(* IEC 61131-3 sources: TetherPLC/tests/compat (part 3) *)

(* ---- tc2_ncfifoaxes_case.st ---- *)
PROGRAM Tc2NciFifoCase
VAR
    mask   AT %QD0 : DINT;
    st     : INT;
    prevSt : INT;
    cur    : INT;
    pulse  : BOOL;
    ax     : FB_MotionAxis;
    axM    : UDINT;
    axS    : UDINT;
    pwrM   : MC_Power;
    pwrS   : MC_Power;
    integ1 : FiFoGroupIntegrate;
    integ2 : FiFoGroupIntegrate;
    dim    : FiFoGetDimension;
    wr     : FiFoWrite;
    owr    : FiFoOverwrite;
    ovr    : FiFoSetChannelOverride;
    start  : FiFoStart;
    dis    : FiFoGroupDisintegrate;
    mon    : FB_Fifo;
    dim2   : FiFoGetDimension;
    rpM    : MC_ReadActualPosition;
    rpS    : MC_ReadActualPosition;
    data   : ARRAY[0..255] OF LREAL;
    k      : UDINT;
    enSig  : BOOL;
    finishedSeen : BOOL;
    seqOk  : BOOL;
    seqOk2 : BOOL;
    posOk1 : BOOL;
    posOk2 : BOOL;
    startEx : BOOL;
END_VAR

// Stage machine: one stage per scan via the cur snapshot.
cur := st;
IF cur <> prevSt THEN pulse := TRUE; ELSE pulse := FALSE; END_IF;
prevSt := cur;

// Channel monitor: status+poll every scan. In-process backends
// consume one queued row per poll; the IO backend consumes rows on
// the mc.time drive clock (poll is a no-op there).
mon.OP := 6;
mon.CHAN := 0;
mon();

enSig := (st >= 1) AND (st <= 40);
// FiFoStart is invoked every scan so its Execute edge tracking stays
// live across the two run stages.
startEx := pulse AND ((cur = 6) OR (cur = 10));
start(bExecute := startEx, iChannelId := 0, tTimeout := T#1S);
pwrM(Enable := enSig, Enable_Positive := TRUE, Enable_Negative := TRUE,
    Axis := axM);
pwrS(Enable := enSig, Enable_Positive := TRUE, Enable_Negative := TRUE,
    Axis := axS);
rpM(Enable := TRUE, Axis := axM);
rpS(Enable := TRUE, Axis := axS);

IF cur = 0 THEN
    ax.UNITS_PER_REV := 1000;
    ax.MAX_VEL := 2000;
    ax.MAX_ACCEL := 8000;
    ax.MAX_DECEL := 8000;
    ax.POS_MIN := -200000;
    ax.POS_MAX := 200000;
    ax.HOME_OFFSET := 0;
    ax.FOLLOW_WINDOW := 3;
    ax.FLAGS := 1;
    ax.OP := 1; ax();
    IF ax.AXIS <> 0 THEN axM := ax.AXIS; END_IF;
    ax.OP := 1; ax();
    IF ax.AXIS <> 0 THEN axS := ax.AXIS; END_IF;
    IF axM <> 0 AND axS <> 0 THEN
        mask := mask + 1;                       // bit0: two axes
        st := 1;
    END_IF;
ELSIF cur = 1 THEN
    IF pwrM.Status AND pwrS.Status THEN
        mask := mask + 2;                       // bit1: powered
        st := 2;
    END_IF;
ELSIF cur = 2 THEN
    integ1(bExecute := pulse, iChannelId := 0, iAxisId := axM,
           iGroupPosition := 1, tTimeout := T#1S);
    integ2(bExecute := pulse, iChannelId := 0, iAxisId := axS,
           iGroupPosition := 2, tTimeout := T#1S);
    IF pulse AND NOT integ1.bError AND NOT integ2.bError THEN
        mask := mask + 4;                       // bit2: integrated
        st := 3;
    END_IF;
ELSIF cur = 3 THEN
    dim(bExecute := pulse, iChannelId := 0, tTimeout := T#1S);
    IF dim.bError = FALSE THEN
        IF dim.iAxes = 2 AND dim.iMaxRows >= 100 THEN
            mask := mask + 8;                   // bit3: dimension
            st := 4;
        END_IF;
    END_IF;
ELSIF cur = 4 THEN
    // two rows x two axes: [100,200] then [300,400]
    data[0] := 100.0; data[1] := 200.0;
    data[8] := 300.0; data[9] := 400.0;
    wr(bExecute := pulse, iChannelId := 0,
       AdrDataArray := data, iRowsToWrite := 2, tTimeout := T#1S);
    IF pulse AND NOT wr.bError THEN
        mask := mask + 16;                      // bit4: write
        st := 5;
    END_IF;
ELSIF cur = 5 THEN
    ovr(bExecute := pulse, iChannelId := 0, iOverride := 150,
        tTimeout := T#1S);
    IF pulse AND NOT ovr.bError THEN
        mask := mask + 32;                      // bit5: override
        st := 6;
    END_IF;
ELSIF cur = 6 THEN
    IF pulse AND NOT start.bError THEN
        mask := mask + 64;                      // bit6: start
        st := 7;
    END_IF;
ELSIF cur = 7 THEN
    // wait for the channel to drain (state 2 = finished)
    IF mon.STATE = 2 THEN
        IF mon.SEQ = 2 THEN
            seqOk := TRUE;
        END_IF;
        finishedSeen := TRUE;
        st := 8;
    END_IF;
ELSIF cur = 8 THEN
    // positions should have snapped/tracked to the last row
    IF rpM.Valid AND rpS.Valid THEN
        IF DINT_TO_LREAL(rpM.Position) >= 295.0 AND
           DINT_TO_LREAL(rpS.Position) >= 395.0 THEN
            posOk1 := TRUE;
        END_IF;
    END_IF;
    IF posOk1 THEN
        mask := mask + 128;                     // bit7: row positions
        st := 9;
    END_IF;
ELSIF cur = 9 THEN
    // overwrite the queue with a single row [500,600] and rerun
    FOR k := 0 TO 255 DO data[k] := 0.0; END_FOR;
    data[0] := 500.0; data[1] := 600.0;
    owr(bExecute := pulse, iChannelId := 0,
        AdrDataArray := data, iRowsToWrite := 1, tTimeout := T#1S);
    IF pulse AND NOT owr.bError THEN
        mask := mask + 256;                     // bit8: overwrite
        st := 10;
    END_IF;
ELSIF cur = 10 THEN
    IF pulse AND NOT start.bError THEN
        st := 11;
    END_IF;
ELSIF cur = 11 THEN
    IF mon.STATE = 2 THEN
        IF mon.SEQ = 1 THEN seqOk2 := TRUE; END_IF;
        st := 12;
    END_IF;
ELSIF cur = 12 THEN
    IF rpM.Valid AND rpS.Valid THEN
        IF DINT_TO_LREAL(rpM.Position) >= 495.0 AND
           DINT_TO_LREAL(rpS.Position) >= 595.0 THEN
            posOk2 := TRUE;
        END_IF;
    END_IF;
    IF posOk2 THEN
        mask := mask + 512;                     // bit9: overwrite pos
        st := 13;
    END_IF;
ELSIF cur = 13 THEN
    dis(bExecute := pulse, iChannelId := 0, tTimeout := T#1S);
    IF pulse AND NOT dis.bError THEN
        dim2(bExecute := pulse, iChannelId := 0, tTimeout := T#1S);
        IF dim2.iAxes = 0 THEN
            mask := mask + 1024;                // bit10: disintegrate
            st := 14;
        END_IF;
    END_IF;
ELSIF cur = 14 THEN
    // final: fold run flags into spare bits (one-shot stage)
    IF seqOk AND seqOk2 THEN mask := mask + 2048; END_IF; // bit11
    IF posOk1 THEN mask := mask + 4096; END_IF;           // bit12
    IF posOk2 THEN mask := mask + 8192; END_IF;           // bit13
    st := 15;
ELSIF cur = 15 THEN
    // hold; expect written at final step
END_IF;
END_PROGRAM

(* ---- tc2_nci_case.st ---- *)
PROGRAM Tc2NciCase
VAR
    mask   AT %QD0 : DINT;
    st     : INT;
    prevSt : INT;
    pulse  : BOOL;
    ax     : FB_MotionAxis;
    axX     : UDINT;
    axY     : UDINT;
    axZ     : UDINT;
    pX     : MC_Power;
    pY     : MC_Power;
    pZ     : MC_Power;
    ln     : FB_NciLine;
    estp   : FB_NciEStop;
    rX     : MC_ReadActualPosition;
    rY     : MC_ReadActualPosition;
    rZ     : MC_ReadActualPosition;
    enSig  : BOOL;
    lnEx   : BOOL;
    estpEx : BOOL;
    lnX    : DINT;
    lnY    : DINT;
    lnZ    : DINT;
END_VAR

// Create the three group axes once.
IF st = 0 THEN
    ax.UNITS_PER_REV := 1000;
    ax.MAX_VEL := 200000;
    ax.MAX_ACCEL := 800000;
    ax.MAX_DECEL := 800000;
    ax.POS_MIN := -2000000;
    ax.POS_MAX := 2000000;
    ax.FLAGS := 1;
    ax.OP := 1; ax();
    IF ax.AXIS <> 0 THEN axX := ax.AXIS; END_IF;
    ax.OP := 1; ax();
    IF ax.AXIS <> 0 THEN axY := ax.AXIS; END_IF;
    ax.OP := 1; ax();
    IF ax.AXIS <> 0 THEN axZ := ax.AXIS; END_IF;
    IF axX <> 0 AND axY <> 0 AND axZ <> 0 THEN
        mask := mask + 1;                       // bit0: 3 axes
    END_IF;
    st := 1;
    prevSt := 0;
END_IF;

IF st <> prevSt THEN pulse := TRUE; ELSE pulse := FALSE; END_IF;
prevSt := st;

enSig  := (st >= 1) AND (st <= 5);
lnEx   := (st = 2) OR (st = 4);    // move1 target, move2 home
estpEx := pulse AND (st = 6);
IF st <= 3 THEN
    lnX := 1000; lnY := 600; lnZ := 300;   // first segment
ELSE
    lnX := 0;    lnY := 0;   lnZ := 0;     // return to origin
END_IF;

pX(Enable := enSig, Enable_Positive := TRUE, Enable_Negative := TRUE,
   Axis := axX);
pY(Enable := enSig, Enable_Positive := TRUE, Enable_Negative := TRUE,
   Axis := axY);
pZ(Enable := enSig, Enable_Positive := TRUE, Enable_Negative := TRUE,
   Axis := axZ);
ln(Execute := lnEx, PosX := lnX, PosY := lnY, PosZ := lnZ,
   Velocity := 2000, CycleUs := 10000,
   AxisX := axX, AxisY := axY, AxisZ := axZ);
estp(Execute := estpEx, AxisX := axX, AxisY := axY, AxisZ := axZ);
rX(Enable := TRUE, Axis := axX);
rY(Enable := TRUE, Axis := axY);
rZ(Enable := TRUE, Axis := axZ);

IF st = 1 THEN
    IF pX.Status AND pY.Status AND pZ.Status THEN
        mask := mask + 2;                    // bit1: group powered
        st := 2;
    END_IF;
ELSIF st = 2 THEN
    // coordinated linear move to (1000,600,300)
    IF ln.Done THEN
        mask := mask + 4;                    // bit2: move1 done
        st := 3;
    END_IF;
ELSIF st = 3 THEN
    // every axis arrived at its target coordinate (CSP == commanded).
    // the actual position lags the streamed target by a scan or two
    // depending on the backend, so wait for it to converge before
    // asserting the endpoint bits and moving on.
    IF rX.Position = 1000 AND rY.Position = 600 AND
       rZ.Position = 300 THEN
        mask := mask + 8;                    // bit3: endpoints hit
        // path length = sqrt(1e6+3.6e5+9e4)=sqrt(1.45e6)=1204.16
        IF ln.PathLen >= 1200 AND ln.PathLen <= 1210 THEN
            mask := mask + 16;               // bit4: path length
        END_IF;
        st := 4;
    END_IF;
ELSIF st = 4 THEN
    // second coordinated move back to the origin
    IF ln.Done THEN
        mask := mask + 32;                   // bit5: move2 done
        st := 5;
    END_IF;
ELSIF st = 5 THEN
    // wait for the positions to converge on the origin (same
    // backend-lag reasoning as st=3)
    IF rX.Position = 0 AND rY.Position = 0 AND
       rZ.Position = 0 THEN
        mask := mask + 64;                   // bit6: back at origin
        st := 6;
    END_IF;
ELSIF st = 6 THEN
    // group E-stop removes power from all three axes
    IF estp.Status THEN
        mask := mask + 128;                  // bit7: all disabled
        st := 7;
    END_IF;
END_IF;

END_PROGRAM

(* ---- tc2_nci_gcode_case.st ---- *)
PROGRAM Tc2NciGcodeCase
VAR
    mask   AT %QD0 : DINT;
    st     : INT;
    prevSt : INT;
    ldt    : FB_ItpLoadText;
    ldf    : FB_ItpLoadProg;
    ss     : FB_ItpStartStop;
    rst    : FB_ItpReset;
    sts    : FB_ItpStatus;
    ldtEx  : BOOL;
    ldfEx  : BOOL;
    stStart : BOOL;
    stStop : BOOL;
    rsEx   : BOOL;
    waitN  : INT;
    fwA    : FB_ItpFiFoWrite;
    fwB    : FB_ItpFiFoWrite;
    cnf    : FB_ItpConfirmHsk;
    rpw    : FB_ItpWriteRParam;
    rpr    : FB_ItpReadRParam;
    zs     : FB_ItpZeroShift;
    fwAEx  : BOOL;
    fwBEx  : BOOL;
    cnfEx  : BOOL;
    rpwEx  : BOOL;
    rprEx  : BOOL;
    zsEx   : BOOL;
    rpDone : BOOL;
    m8Seen : BOOL;
END_VAR

// The 7-block program lives on the server host (the shell script
// writes /tmp/tplc_nci_case.g before the sim runs); inline text is
// exercised with a tiny two-block program.
IF st = 0 THEN
    mask := 0;
    st := 1;
END_IF;

IF st <> prevSt THEN waitN := 0; END_IF;
prevSt := st;
waitN := waitN + 1;

ldtEx   := (st = 1) AND (waitN = 2);
ldfEx   := (st = 4) AND (waitN = 2);
stStart := ((st = 6) OR (st = 14) OR (st = 19)) AND (waitN = 2);
stStop  := (st = 10) AND (waitN = 2);
rsEx    := (st = 3) OR (st = 11) OR (st = 16) OR (st = 21);
rsEx    := rsEx AND (waitN = 2);
fwAEx   := (st = 13) AND (waitN = 2);
fwBEx   := (st = 13) AND (waitN = 3);
rpwEx   := (st = 18) AND (waitN = 2);
rprEx   := (st = 18) AND (waitN = 4);
zsEx    := (st = 18) AND (waitN = 6);
cnfEx   := (st = 19) AND (sts.MFunc = 8);

sts(ChanId := 0);
ldt(Execute := ldtEx, ChanId := 0,
    ProgText := 'G1 X1 F600$NM30$N');
ldf(Execute := ldfEx, ChanId := 0,
    PathName := '/tmp/tplc_nci_case.g');
ss(Start := stStart, Stop := stStop, ChanId := 0);
rst(Execute := rsEx, ChanId := 0);
fwA(Execute := fwAEx, ChanId := 0, Block := 'G1 X2 F600');
fwB(Execute := fwBEx, ChanId := 0, Block := 'G1 X0 F600');
cnf(Execute := cnfEx, ChanId := 0);
rpw(Execute := rpwEx, ChanId := 0, Index := 100, Value := 42.5);
rpr(Execute := rprEx, ChanId := 0, Index := 100);
zs(Execute := zsEx, ChanId := 0, OffX := 5.0, OffY := 0.0, OffZ := 0.0);

IF st = 1 THEN
    // inline text upload accepted
    IF ldt.Done THEN
        mask := mask + 1;                    // bit0: text upload ok
        st := 2;
    ELSIF ldt.Error THEN
        st := 90;
    END_IF;
ELSIF st = 2 THEN
    // compiled: READY (state 1) with 2 blocks
    IF sts.Valid AND (sts.State = 1) THEN
        mask := mask + 2;                    // bit1: ready
        IF sts.Total = 2 THEN
            mask := mask + 4;                // bit2: 2 blocks
        END_IF;
        st := 3;
    ELSIF sts.Valid AND (sts.State = 5) THEN
        st := 91;
    END_IF;
ELSIF st = 3 THEN
    // reset back to IDLE before the file load
    IF rst.Done THEN
        mask := mask + 8;                    // bit3: reset ok
        st := 4;
    ELSIF rst.Error THEN
        st := 92;
    END_IF;
ELSIF st = 4 THEN
    // file load accepted
    IF ldf.Done THEN
        mask := mask + 16;                   // bit4: file load ok
        st := 5;
    ELSIF ldf.Error THEN
        st := 93;
    END_IF;
ELSIF st = 5 THEN
    // file compiled: READY with 7 blocks
    IF sts.Valid AND (sts.State = 1) THEN
        mask := mask + 32;                   // bit5: ready
        IF sts.Total = 7 THEN
            mask := mask + 64;               // bit6: 7 blocks
        END_IF;
        st := 6;
    ELSIF sts.Valid AND (sts.State = 5) THEN
        st := 94;
    END_IF;
ELSIF st = 6 THEN
    IF ss.Done THEN
        mask := mask + 128;                  // bit7: run accepted
        st := 7;
    ELSIF ss.Error THEN
        st := 95;
    END_IF;
ELSIF st = 7 THEN
    // running: mid-program block reached or raced to finish
    IF sts.Valid AND (sts.State = 2) AND (sts.Line >= 3) THEN
        mask := mask + 256;                  // bit8: mid-program
        st := 8;
    ELSIF sts.Valid AND (sts.State = 4) THEN
        st := 8;
    END_IF;
ELSIF st = 8 THEN
    IF sts.Valid AND (sts.State = 4) THEN
        mask := mask + 512;                  // bit9: finished
        st := 9;
    ELSIF sts.Valid AND (sts.State = 5) THEN
        st := 96;
    END_IF;
ELSIF st = 9 THEN
    // planned duration ~4.1s at the given feeds
    IF sts.DurationMs >= 3500 AND sts.DurationMs <= 5000 THEN
        mask := mask + 1024;                 // bit10: duration sane
    END_IF;
    st := 10;
ELSIF st = 10 THEN
    // permissive stop after finish
    IF ss.Done THEN
        mask := mask + 2048;                 // bit11: stop ok
        st := 11;
    ELSIF ss.Error THEN
        st := 97;
    END_IF;
ELSIF st = 11 THEN
    IF rst.Done THEN
        mask := mask + 4096;                 // bit12: reset ok
        st := 12;
    ELSIF rst.Error THEN
        st := 98;
    END_IF;
ELSIF st = 12 THEN
    // reset returns the channel to IDLE with no program
    IF sts.Valid AND (sts.State = 0) AND (sts.Total = 0) THEN
        mask := mask + 8192;                 // bit13: idle cleared
        st := 13;
    END_IF;
ELSIF st = 13 THEN
    // two FIFO blocks queued (Done pulses are per-scan; the queue
    // depth is the real check)
    IF sts.Valid AND sts.FifoLen = 2 THEN
        mask := mask + 16384;                // bit14: fifo queued
        st := 14;
    END_IF;
ELSIF st = 14 THEN
    // run the FIFO-only program from idle (stStart pulses above)
    IF ss.Done THEN
        st := 15;
    END_IF;
ELSIF st = 15 THEN
    // both FIFO entries consumed, channel finished
    IF sts.Valid AND (sts.State = 4) AND (sts.FifoSeq = 2) THEN
        mask := mask + 32768;                // bit15: fifo chained
        st := 16;
    END_IF;
ELSIF st = 16 THEN
    IF rst.Done THEN
        mask := mask + 65536;                // bit16: reset ok
        st := 17;
    END_IF;
ELSIF st = 17 THEN
    // M-func program: M8 pauses the channel with pending code
    ldt(Execute := TRUE, ChanId := 0,
        ProgText := 'G21 G90$NG1 X5 F600$NM8$NG1 X10$NM30$N');
    IF ldt.Done THEN
        st := 18;
    END_IF;
ELSIF st = 18 THEN
    // R-param roundtrip + zero-shift write in the same wait window
    IF rpw.Done THEN mask := mask + 131072; END_IF;   // bit17: rp write
    IF rpr.Done AND (rpr.Value > 42.0) AND (rpr.Value < 43.0) THEN
        mask := mask + 262144;                        // bit18: rp read
        rpDone := TRUE;
    END_IF;
    IF zs.Done THEN mask := mask + 524288; END_IF;    // bit19: zshift
    IF (mask AND 917504) = 917504 THEN
        st := 19;
    END_IF;
ELSIF st = 19 THEN
    // run the M-func program; it pauses on M8 (stStart pulses above)
    IF sts.Valid AND (sts.MFunc = 8) AND NOT m8Seen THEN
        mask := mask + 1048576;                // bit20: M8 pending
        m8Seen := TRUE;
    END_IF;
    IF sts.Valid AND (sts.State = 4) AND
       (sts.MFunc = 0) THEN
        mask := mask + 2097152;                // bit21: resumed+done
        st := 20;
    END_IF;
ELSIF st = 20 THEN
    st := 21;
ELSIF st = 21 THEN
    IF rst.Done THEN
        mask := mask + 4194304;                // bit22: reset ok
        st := 22;
    END_IF;
END_IF;

END_PROGRAM

(* ---- tc2_nckin_case.st ---- *)
PROGRAM Tc2NcKinCase
VAR
    mask   AT %QD0 : DINT;
    st     : INT;
    prevSt : INT;
    cur    : INT;
    pulse  : BOOL;
    cfgA   : FB_Kin;
    cfgB   : FB_Kin;
    grp0   : FB_KinConfigGroup;
    grp1   : FB_KinConfigGroup;
    opst   : F_KinGetChnOperationState;
    ids0   : F_KinGetAcsMcsAxisIds;
    ids1   : F_KinGetAcsMcsAxisIds;
    xf     : FB_KinCalcTrafo;
    xb     : FB_KinCalcTrafo;
    xf5    : FB_KinCalcTrafo;
    xf99   : FB_KinCalcTrafo;
    mf     : FB_KinCalcMultiTrafo;
    mb     : FB_KinCalcMultiTrafo;
    mf2    : FB_KinCalcMultiTrafo;
    unl    : FB_KinUnlockTrafoParam;
    lck    : FB_KinLockTrafoParam;
    rotP   : FB_KinPresetRotation;
    extR   : FB_KinExtendedRotationRange;
    rst    : FB_KinResetGroup;
    chk    : FB_KinCheckActualStatus;
    kinSt  : UDINT;
    inA    : ARRAY[0..7] OF LREAL;
    outA   : ARRAY[0..7] OF LREAL;
    ms     : UDINT;
    me     : UDINT;
    inM    : ARRAY[0..7] OF LREAL;
    outM   : ARRAY[0..15] OF LREAL;
    inM2   : ARRAY[0..7] OF LREAL;
    outM2  : ARRAY[0..15] OF LREAL;
    acsArr : ARRAY[0..7] OF UDINT;
    mcsArr : ARRAY[0..7] OF UDINT;
    acsEmp : ARRAY[0..7] OF UDINT;
    mcsEmp : ARRAY[0..7] OF UDINT;
    rotArr : ARRAY[0..2] OF LREAL;
    tgt    : ARRAY[0..7] OF LREAL;
    jnt    : ARRAY[0..7] OF LREAL;
    posA   : ARRAY[0..7] OF LREAL;
    posB   : ARRAY[0..7] OF LREAL;
    tolA   : ARRAY[0..7] OF LREAL;
    tolOk1 : BOOL;
    tolOk2 : BOOL;
    started : BOOL;
    i      : UDINT;
END_VAR

cur := st;
/* pulse on stage entry; the very first scan counts too (prevSt
   would otherwise equal cur=0 and swallow the st0 edge). */
pulse := (cur <> prevSt) OR NOT started;
started := TRUE;
prevSt := cur;

// Persistent inputs for the edge-triggered wrappers (called every
// scan so their internal Execute edge tracking stays live).
FOR i := 0 TO 7 DO
    acsArr[i] := 0;
    mcsArr[i] := 0;
    inA[i] := 0.0;
    outA[i] := 0.0;
END_FOR;
acsArr[0] := 1; acsArr[1] := 2;
mcsArr[0] := 3; mcsArr[1] := 4; mcsArr[2] := 5;
rotArr[0] := 0.1; rotArr[1] := 0.2; rotArr[2] := 0.3;
kinSt := 0;

// st0: configure obj0 = planar2d (L1=L2=0.5), obj1 = serial6 UR5
grp0(bExecute := FALSE, bCartesianMode := FALSE, oidTrafo := 0,
     nItpChannelId := 0, AcsAxis := acsArr, McsAxis := mcsArr);
grp1(bExecute := FALSE, bCartesianMode := FALSE, oidTrafo := 1,
     nItpChannelId := 0, AcsAxis := acsEmp, McsAxis := mcsEmp);
IF cur = 0 THEN
    IF pulse THEN
        cfgA.OBJ := 0; cfgA.OP := 1; cfgA.TYPEIN := 1;
        cfgA.PRESET := 0; cfgA.NCFG := 2;
        cfgA.CFG[0] := 0.5; cfgA.CFG[1] := 0.5;
        cfgA();
        cfgB.OBJ := 1; cfgB.OP := 1; cfgB.TYPEIN := 4;
        cfgB.PRESET := 0; cfgB.NCFG := 0;
        cfgB();
        IF cfgA.STATUS = 0 AND cfgB.STATUS = 0 THEN
            mask := mask + 1;                   // bit0: configure
        END_IF;
    END_IF;
    st := 1;
// st1: bind axes + channel on both objects
ELSIF cur = 1 THEN
    grp0(bExecute := pulse, bCartesianMode := FALSE, oidTrafo := 0,
         nItpChannelId := 7, AcsAxis := acsArr, McsAxis := mcsArr);
    grp1(bExecute := pulse, bCartesianMode := FALSE, oidTrafo := 1,
         nItpChannelId := 0, AcsAxis := acsEmp, McsAxis := mcsEmp);
    IF pulse AND NOT grp0.bError AND NOT grp1.bError THEN
        mask := mask + 2;                       // bit1: config group
    END_IF;
    st := 2;
// st2: op state + axis list readback
ELSIF cur = 2 THEN
    opst(oidTrafo := 0);
    ids0(oidTrafo := 0);
    ids1(oidTrafo := 1);
    IF opst.OpState = 1 AND opst.ErrorId = 0 AND
       ids0.ErrorId = 0 AND ids0.NAcs = 2 AND ids0.NMcs = 3 AND
       ids0.AcsAxis[0] = 1 AND ids0.AcsAxis[1] = 2 AND
       ids0.McsAxis[0] = 3 AND ids0.McsAxis[2] = 5 AND
       ids1.NAcs = 0 THEN
        mask := mask + 4;                       // bit2: status/axes
    END_IF;
    st := 3;
// st3: forward transform planar2d q={0.3,0.4}
ELSIF cur = 3 THEN
    inA[0] := 0.3; inA[1] := 0.4;
    xf(bExecute := pulse, bForward := TRUE, oidTrafo := 0,
       AxesPosIn := inA, AxesPosOut := outA,
       MetaState := ms, MetaError := me);
    IF pulse AND NOT xf.bError AND
       ABS(outA[0] - 0.8601) < 0.01 AND
       ABS(outA[1] - 0.4699) < 0.01 AND
       ABS(outA[2]) < 0.001 THEN
        mask := mask + 8;                       // bit3: forward
    END_IF;
    st := 4;
// st4: backward IK to the same target, seeded near the solution
ELSIF cur = 4 THEN
    inA[0] := 0.8601; inA[1] := 0.4699; inA[2] := 0.0;
    inA[3] := 0.3; inA[4] := 0.4;
    xb(bExecute := pulse, bForward := FALSE, oidTrafo := 0,
       AxesPosIn := inA, AxesPosOut := outA,
       MetaState := ms, MetaError := me);
    IF pulse AND NOT xb.bError AND me = 0 AND
       ABS(outA[0] - 0.3) < 0.05 AND
       ABS(outA[1] - 0.4) < 0.05 THEN
        mask := mask + 16;                      // bit4: inverse IK
    END_IF;
    st := 5;
// st5: CalcMultiTrafo forward on serial6 UR5, q={0.1..0.6}
ELSIF cur = 5 THEN
    inM[0] := 0.1; inM[1] := 0.2; inM[2] := 0.3;
    inM[3] := 0.4; inM[4] := 0.5; inM[5] := 0.6;
    mf(bExecute := pulse, bForward := TRUE, oidTrafo := 1,
       nSizeIn := 6, nSizeOut := 16,
       InData := inM, OutData := outM);
    IF pulse AND NOT mf.bError THEN
        tgt[0] := outM[0]; tgt[1] := outM[1]; tgt[2] := outM[2];
        mask := mask + 32;                      // bit5: multi fwd
    END_IF;
    st := 6;
// st6: CalcMultiTrafo backward IK on the serial6 target
ELSIF cur = 6 THEN
    inM2[0] := tgt[0]; inM2[1] := tgt[1]; inM2[2] := tgt[2];
    inM2[3] := 0.1; inM2[4] := 0.2; inM2[5] := 0.3;
    mb(bExecute := pulse, bForward := FALSE, oidTrafo := 1,
       nSizeIn := 7, nSizeOut := 16,
       InData := inM2, OutData := outM2);
    IF pulse AND NOT mb.bError THEN
        FOR i := 0 TO 5 DO jnt[i] := outM2[i]; END_FOR;
        mask := mask + 64;                      // bit6: multi inv
    END_IF;
    st := 7;
// st7: forward again with the IK joints; pose must match target
ELSIF cur = 7 THEN
    FOR i := 0 TO 5 DO inM[i] := jnt[i]; END_FOR;
    mf2(bExecute := pulse, bForward := TRUE, oidTrafo := 1,
        nSizeIn := 6, nSizeOut := 16,
        InData := inM, OutData := outM2);
    IF pulse AND NOT mf2.bError AND
       ABS(outM2[0] - tgt[0]) < 0.001 AND
       ABS(outM2[1] - tgt[1]) < 0.001 AND
       ABS(outM2[2] - tgt[2]) < 0.001 THEN
        mask := mask + 128;                     // bit7: ik roundtrip
    END_IF;
    st := 8;
// st8: preset rotation A = {0.1,0.2,0.3}
ELSIF cur = 8 THEN
    rotP(bExecute := pulse, oidTrafo := 0, Rotation := rotArr);
    st := 9;
// st9: extended range saves A (edge), then preset B overwrites
ELSIF cur = 9 THEN
    extR(bExecute := TRUE, oidTrafo := 0);
    rotArr[0] := 0.9; rotArr[1] := 0.8; rotArr[2] := 0.7;
    rotP(bExecute := pulse, oidTrafo := 0, Rotation := rotArr);
    st := 10;
// st10: hold extended (no edge yet)
ELSIF cur = 10 THEN
    extR(bExecute := TRUE, oidTrafo := 0);
    st := 11;
// st11: release -> restore A
ELSIF cur = 11 THEN
    extR(bExecute := FALSE, oidTrafo := 0);
    st := 12;
// st12: rotation state must be A again
ELSIF cur = 12 THEN
    cfgA.OBJ := 0; cfgA.OP := 7; cfgA.ROP := 0; cfgA();
    IF ABS(cfgA.ROT[0] - 0.1) < 0.0001 AND
       ABS(cfgA.ROT[1] - 0.2) < 0.0001 AND
       ABS(cfgA.ROT[2] - 0.3) < 0.0001 THEN
        mask := mask + 256;                     // bit8: rotation
    END_IF;
    st := 13;
// st13: reset group on obj0
ELSIF cur = 13 THEN
    rst(bExecute := pulse, oidTrafo := 0, nItpChannelId := 0);
    st := 14;
// st14: channel op state now idle; tolerance function checks
ELSIF cur = 14 THEN
    chk(bExecute := pulse, oidTrafo := 0, eKinStatus := kinSt);
    FOR i := 0 TO 7 DO
        posA[i] := 0.0; posB[i] := 0.0; tolA[i] := 0.0;
    END_FOR;
    posA[0] := 1.0; posA[1] := 2.0; posA[2] := 3.0;
    posB[0] := 1.0000001; posB[1] := 2.0; posB[2] := 3.0;
    tolA[0] := 0.001; tolA[1] := 0.001; tolA[2] := 0.001;
    tolOk1 := F_KinAxesInTolerance(posA, posB, tolA);
    posB[0] := 2.0;
    tolOk2 := F_KinAxesInTolerance(posA, posB, tolA);
    IF kinSt = 0 AND tolOk1 AND NOT tolOk2 THEN
        mask := mask + 512;                     // bit9: reset+tolerance
    END_IF;
    st := 15;
// st15: transform on an unconfigured object -> MetaError = 1
ELSIF cur = 15 THEN
    xf5(bExecute := pulse, bForward := TRUE, oidTrafo := 5,
        AxesPosIn := inA, AxesPosOut := outA,
        MetaState := ms, MetaError := me);
    IF pulse AND NOT xf5.bError AND me = 1 THEN
        mask := mask + 1024;                    // bit10: no-model err
    END_IF;
    st := 16;
// st16: out-of-range object id -> transport-level error
ELSIF cur = 16 THEN
    xf99(bExecute := pulse, bForward := TRUE, oidTrafo := 99,
         AxesPosIn := inA, AxesPosOut := outA,
         MetaState := ms, MetaError := me);
    IF pulse AND xf99.bError THEN
        mask := mask + 2048;                    // bit11: bad obj
    END_IF;
    st := 17;
// st17: parameter lock — unlock, reconfigure OK, lock, configure
// must be rejected with E_LOCKED (-4)
ELSIF cur = 17 THEN
    IF pulse THEN
        unl(bExecute := TRUE, oidTrafo := 0);
        cfgA.OBJ := 0; cfgA.OP := 1; cfgA.TYPEIN := 1;
        cfgA.PRESET := 0; cfgA.NCFG := 0; cfgA();
        IF unl.bError = FALSE AND cfgA.STATUS = 0 THEN
            lck(bExecute := TRUE, oidTrafo := 0);
            cfgA.OBJ := 0; cfgA.OP := 1; cfgA.TYPEIN := 3;
            cfgA.PRESET := 0; cfgA.NCFG := 0; cfgA();
            IF lck.bError = FALSE AND cfgA.STATUS = -4 THEN
                mask := mask + 4096;            // bit12: lock
            END_IF;
        END_IF;
    END_IF;
    st := 18;
ELSIF cur = 18 THEN
    // hold; expect written at final step
END_IF;
END_PROGRAM

(* ---- tc2_ocpp_case.st ---- *)
// tc2_ocpp_case.st — OCPP-J client e2e over the python CSMS fake.
// WS upgrade, OCPP call -> echoed result, disconnect.
PROGRAM tc2_ocpp_case
VAR
    con : FB_OcppConnect;
    dis : FB_OcppDisconnect;
    cal : FB_OcppCall;
    rx  : FB_OcppReceive;
    st : INT;
    waitN : INT;
    mask AT %QD0 : UDINT;
    hdl : UDINT;
END_VAR
    IF st = 0 THEN
        mask := 0;
        con.Execute := TRUE;
        con.Host := '127.0.0.1';
        con.Port := 11890;
        con.Path := '/ocpp';
        con.ChargePointId := 'CP001';
        st := 1;
    END_IF;

    IF st = 1 THEN
        IF con.Done THEN
            hdl := con.ConnectionHdl;
            con.Execute := FALSE;
            mask := mask + 1;         // bit0: ws session up
            cal.Execute := TRUE;
            cal.ConnectionHdl := hdl;
            cal.MessageId := 'boot-1';
            cal.ActName := 'BootNotification';
            cal.Payload := '{"chargePointVendor":"Tether","chargePointModel":"TPLC"}';
            st := 2;
        END_IF;
        IF con.Error THEN mask := 16#DEAD; st := 99; END_IF;
    END_IF;

    IF st = 2 THEN
        IF cal.Done THEN
            mask := mask + 2;         // bit1: call sent
            cal.Execute := FALSE;
            rx.Execute := TRUE;
            rx.ConnectionHdl := hdl;
            st := 3;
        END_IF;
        IF cal.Error THEN mask := 16#DEAD; st := 99; END_IF;
    END_IF;

    // poll for the CSMS fake's echoed result
    IF st = 3 THEN
        waitN := waitN + 1;
        IF rx.Message THEN
            IF rx.MessageType = 3 THEN
                mask := mask + 4;     // bit2: result landed
            END_IF;
            rx.Execute := FALSE;
            dis.Execute := TRUE;
            dis.ConnectionHdl := hdl;
            st := 4;
        END_IF;
        IF rx.Error THEN mask := 16#DEAD; st := 99; END_IF;
        IF waitN > 40 THEN
            rx.Execute := FALSE;
            dis.Execute := TRUE;
            dis.ConnectionHdl := hdl;
            st := 4;
        END_IF;
    END_IF;

    IF st = 4 THEN
        IF dis.Done THEN
            mask := mask + 8;         // bit3: released
            st := 5;
        END_IF;
        IF dis.Error THEN mask := 16#DEAD; st := 99; END_IF;
    END_IF;

    con(); dis(); cal(); rx();
END_PROGRAM

(* ---- tc2_opcua_case.st ---- *)
// tc2_opcua_case.st — OPC UA client e2e over the open62541 endpoint.
// Connects to the tether_io_motion_server --opcua listener, reads
// nc.state (U8), writes nc.scale=500.0 (F64), reads it back, then
// disconnects. The final mask lands in out 0.
PROGRAM tc2_opcua_case
VAR
    con : FB_UA_Connect;
    dis : FB_UA_Disconnect;
    sta : FB_UA_ConnectGetStatus;
    rd  : FB_UA_Read;
    wr  : FB_UA_Write;
    nsi : FB_UA_GetNamespaceIndex;
    st : INT;
    waitN : INT;
    mask AT %QD0 : UDINT;
    hdl : UDINT;
END_VAR

    // ---- state machine ----
    IF st = 0 THEN
        mask := 0;
        con.Execute := TRUE;
        con.ServerUrl := 'opc.tcp://[::1]:14199';
        st := 1;
    END_IF;

    IF st = 1 THEN
        IF con.Done THEN
            hdl := con.ConnectionHdl;
            con.Execute := FALSE;
            mask := mask + 1;         // bit0: connected
            st := 2;
            waitN := 0;
        END_IF;
        IF con.Error THEN
            mask := 16#DEAD;
            st := 99;
        END_IF;
    END_IF;

    IF st = 2 THEN
        waitN := waitN + 1;
        IF waitN >= 10 THEN
            sta.Execute := TRUE;
            sta.ConnectionHdl := hdl;
            st := 3;
        END_IF;
    END_IF;

    IF st = 3 THEN
        IF sta.Done THEN
            IF sta.ConnectionState = 1 THEN   // TPLC_UA_CONN_OPEN
                mask := mask + 2;             // bit1: session open
                sta.Execute := FALSE;
                rd.Execute := TRUE;
                rd.ConnectionHdl := hdl;
                rd.NodeId := 'ns=2;s=nc.state';
                st := 4;
            END_IF;
        END_IF;
        IF sta.Error THEN
            mask := 16#DEAD;
            st := 99;
        END_IF;
    END_IF;

    IF st = 4 THEN
        IF rd.Done THEN
            IF rd.ValueType = 3 THEN          // U8 maps to U64 family
                mask := mask + 4;             // bit2: nc.state read
            END_IF;
            rd.Execute := FALSE;
            wr.Execute := TRUE;
            wr.ConnectionHdl := hdl;
            wr.NodeId := 'ns=2;s=nc.scale';
            wr.Value := 500.0;
            wr.ValueType := 4;                // F64
            st := 5;
        END_IF;
        IF rd.Error THEN
            mask := 16#DEAD;
            st := 99;
        END_IF;
    END_IF;

    IF st = 5 THEN
        IF wr.Done THEN
            mask := mask + 8;                 // bit3: nc.scale written
            wr.Execute := FALSE;
            rd.Execute := TRUE;
            rd.NodeId := 'ns=2;s=nc.scale';
            st := 6;
        END_IF;
        IF wr.Error THEN
            mask := 16#DEAD;
            st := 99;
        END_IF;
    END_IF;

    IF st = 6 THEN
        IF rd.Done THEN
            IF rd.Value > 499.0 AND rd.Value < 501.0 THEN
                mask := mask + 16;            // bit4: nc.scale==500
            END_IF;
            rd.Execute := FALSE;
            nsi.Execute := TRUE;
            nsi.ConnectionHdl := hdl;
            nsi.NamespaceUri := 'http://tether.io/params';
            st := 7;
        END_IF;
        IF rd.Error THEN
            mask := 16#DEAD;
            st := 99;
        END_IF;
    END_IF;

    IF st = 7 THEN
        IF nsi.Done THEN
            IF nsi.NamespaceIndex = 2 THEN
                mask := mask + 32;            // bit5: ns index 2
            END_IF;
            nsi.Execute := FALSE;
            dis.Execute := TRUE;
            dis.ConnectionHdl := hdl;
            st := 8;
        END_IF;
        IF nsi.Error THEN
            mask := 16#DEAD;
            st := 99;
        END_IF;
    END_IF;

    IF st = 8 THEN
        IF dis.Done THEN
            mask := mask + 64;                // bit6: disconnected
            st := 9;
        END_IF;
        IF dis.Error THEN
            mask := 16#DEAD;
            st := 99;
        END_IF;
    END_IF;

    con(); dis(); sta(); rd(); wr(); nsi();
END_PROGRAM

(* ---- tc2_packml_case.st ---- *)
// tc2_packml_case.st — PackML state machine e2e: Idle -> Start ->
// Execute -> Hold -> Held -> Unhold -> Execute -> Abort -> Aborted
// -> Clear -> Idle.  Command constants per tc2_packml.st header.
PROGRAM tc2_packml_case
VAR
    pml : FB_PackML;
    st : INT;
    waitN : INT;
    mask AT %QD0 : UDINT;
END_VAR
    IF st = 0 THEN
        mask := 0;
        pml.Execute := TRUE;
        pml.Busy := FALSE;
        pml.Command := 0;
        st := 1;
    END_IF;

    // Idle -> Start -> Execute
    IF st = 1 THEN
        IF pml.State = 1 THEN              // Idle
            mask := mask + 1;
            pml.Command := 1;              // Start
            st := 2;
        END_IF;
    END_IF;
    IF st = 2 THEN
        IF pml.State = 3 THEN              // Execute
            mask := mask + 2;
            pml.Command := 4;              // Hold
            st := 3;
        END_IF;
    END_IF;
    // Execute -> Hold -> Held -> Unhold -> Execute
    IF st = 3 THEN
        IF pml.State = 8 THEN              // Held
            mask := mask + 4;
            pml.Command := 5;              // Unhold
            st := 4;
        END_IF;
    END_IF;
    IF st = 4 THEN
        IF pml.State = 3 THEN              // Execute again
            mask := mask + 8;
            pml.Command := 8;              // Abort
            st := 5;
        END_IF;
    END_IF;
    // Execute -> Abort -> Aborted -> Clear -> Idle
    IF st = 5 THEN
        IF pml.State = 14 THEN             // Aborted
            mask := mask + 16;
            pml.Command := 9;              // Clear
            st := 6;
        END_IF;
    END_IF;
    IF st = 6 THEN
        IF pml.State = 1 THEN              // back to Idle
            mask := mask + 32;
            pml.Command := 0;
            st := 7;
        END_IF;
    END_IF;

    pml();
END_PROGRAM

(* ---- tc2_pfwlib_case.st ---- *)
// tc2_pfwlib_case.st — TcTvA alarm-queue e2e: append x2, query,
// deactivate, garbage-collect, clear-pending, clear-signal,
// update-time.  Commands are edge-triggered (nCmd held 0 between);
// ELSIF chain prevents same-scan state cascade.
PROGRAM tc2_pfwlib_case
VAR
    q : FB_TcTvAMsgQueue;
    st : INT;
    mask AT %QD0 : UDINT;
END_VAR
    IF st = 0 THEN
        mask := 0;
        q.nCmd := 0;
        st := 1;
    ELSIF st = 1 THEN
        q.Idx1 := 1; q.Idx2 := 2; q.ErrorId := 100; q.Prio := 3;
        q.Tick := 1000; q.nCmd := 1;
        st := 2;
    ELSIF st = 2 THEN
        q.nCmd := 0;
        IF q.bDone AND q.Count = 1 THEN mask := mask + 1; END_IF;
        st := 3;
    ELSIF st = 3 THEN
        q.Idx1 := 1; q.Idx2 := 2; q.ErrorId := 200; q.Prio := 2;
        q.Tick := 1001; q.nCmd := 1;
        st := 4;
    ELSIF st = 4 THEN
        q.nCmd := 0;
        IF q.bDone AND q.Count = 2 THEN mask := mask + 2; END_IF;
        st := 5;
    ELSIF st = 5 THEN
        // duplicate of A -> reactivates, count stays 2
        q.Idx1 := 1; q.Idx2 := 2; q.ErrorId := 100; q.Prio := 3;
        q.Tick := 1002; q.nCmd := 1;
        st := 6;
    ELSIF st = 6 THEN
        q.nCmd := 0;
        IF q.bDone AND q.Count = 2 THEN mask := mask + 4; END_IF;
        q.QSlot := 0;
        st := 7;
    ELSIF st = 7 THEN
        IF q.QUsed AND q.QActive AND q.QSignaled
           AND q.QIdx1 = 1 AND q.QIdx2 = 2 AND q.QErrorId = 100
           AND q.QPrio = 3 THEN
            mask := mask + 8;
        END_IF;
        st := 8;
    ELSIF st = 8 THEN
        q.Idx1 := 1; q.Idx2 := 2; q.ErrorId := 100; q.Prio := 3;
        q.nCmd := 4;             // deactivate A
        st := 9;
    ELSIF st = 9 THEN
        q.nCmd := 0;
        q.QSlot := 0;
        IF q.bDone AND NOT q.QActive AND q.QUsed THEN
            mask := mask + 16;
        END_IF;
        st := 10;
    ELSIF st = 10 THEN
        q.nCmd := 5;             // garbage collect
        st := 11;
    ELSIF st = 11 THEN
        q.nCmd := 0;
        IF q.bDone AND q.bSignaled AND q.Count = 2 THEN
            mask := mask + 32;
        END_IF;
        st := 12;
    ELSIF st = 12 THEN
        q.Idx1 := 1; q.Idx2 := 2; q.ErrorId := 200; q.Prio := 2;
        q.QSlot := 1;
        q.nCmd := 3;             // clear signal on B
        st := 13;
    ELSIF st = 13 THEN
        q.nCmd := 0;
        IF q.bDone AND NOT q.QSignaled AND q.QActive THEN
            mask := mask + 64;
        END_IF;
        st := 14;
    ELSIF st = 14 THEN
        // clear pending: drop inactive entries with Idx1 in [1..1];
        // A (inactive) removed, B (active) kept -> count 1
        q.IdxFirst := 1; q.IdxLast := 1;
        q.QSlot := 0;
        q.nCmd := 2;
        st := 15;
    ELSIF st = 15 THEN
        q.nCmd := 0;
        IF q.bDone AND q.Count = 1 THEN mask := mask + 128; END_IF;
        st := 16;
    ELSIF st = 16 THEN
        // remaining slot0 is B: active, signal cleared
        IF q.QUsed AND q.QErrorId = 200 AND q.QActive
           AND NOT q.QSignaled THEN
            mask := mask + 256;
        END_IF;
        st := 17;
    ELSIF st = 17 THEN
        q.Tick := 7777; q.nCmd := 6;   // update time
        st := 18;
    ELSIF st = 18 THEN
        q.nCmd := 0;
        IF q.bDone AND q.QTick = 7777 THEN mask := mask + 512; END_IF;
        st := 19;
    ELSIF st = 19 THEN
        q.nCmd := 99;            // unknown command
        st := 20;
    ELSIF st = 20 THEN
        q.nCmd := 0;
        IF q.bError AND q.ErrCode = 16#8002 THEN
            mask := mask + 1024;
        END_IF;
        st := 21;
    END_IF;
    q();
END_PROGRAM

(* ---- tc2_plastic_case.st ---- *)
// tc2_plastic_case.st — Plastic shot-cycle e2e: fill -> pack ->
// hold -> complete with a simulated screw/cavity.
PROGRAM tc2_plastic_case
VAR
    mask AT %QD0 : UDINT;
    shot : FB_PlasticShot;
    screw : LREAL;
    cavity : LREAL;
    st : INT;
    n : INT;
    pSeen : LREAL;
END_VAR
    // One state per scan (ELSIF): outputs read here are the
    // previous call's, inputs written here reach the call below.
    IF st = 0 THEN
        mask := 0;
        screw := 0.0;
        cavity := 0.0;
        n := 0;
        shot.Execute := TRUE;
        shot.StartCycle := FALSE;
        shot.MoldTarget := 80.0;
        shot.FillVel := 40.0;
        shot.CoolTime := 0.3;
        shot.ShotSize := 100.0;
        shot.VpSwitchPos := 20.0;
        shot.CycleTime := 0.1;
        st := 1;
    ELSIF st = 1 THEN
        shot.StartCycle := TRUE;
        st := 2;
    ELSIF st = 2 THEN
        // wait for the fill phase, then release start
        IF shot.Phase = 1 THEN
            mask := mask OR 1;
            shot.StartCycle := FALSE;
            st := 3;
        END_IF;
    ELSIF st = 3 THEN
        // fill: velocity setpoint drives the screw to V/P
        IF shot.VelSetpoint > 0.0 THEN mask := mask OR 2; END_IF;
        shot.ScrewPos := shot.ScrewPos + 4.0;
        IF shot.Phase = 2 THEN
            mask := mask OR 4;
            st := 4;
        END_IF;
    ELSIF st = 4 THEN
        // pack: cavity pressure rises to the pack setpoint
        pSeen := shot.PressureSetpoint;
        IF pSeen > 70.0 THEN mask := mask OR 8; END_IF;
        shot.CavityPressure := 100.0;
        IF shot.Phase = 3 THEN
            mask := mask OR 16;
            st := 5;
        END_IF;
    ELSIF st = 5 THEN
        // complete (start was released in st=2)
        IF shot.CycleFinished THEN
            mask := mask OR 32;
            st := 6;
        END_IF;
    END_IF;

    shot();
END_PROGRAM

(* ---- tc2_pm_case.st ---- *)
// tc2_pm_case.st — PowerMonitoring e2e: V/I sine samples ->
// RMS/P/S/Q/PF/Energy.  The plant feeds a sinusoidal V and a
// in-phase I (PF ~1).
PROGRAM tc2_pm_case
VAR
    pm : FB_PowerMonitor;
    ph : LREAL;   // phase accumulator
    st : INT;
    n : INT;
    mask AT %QD0 : UDINT;
END_VAR
    IF st = 0 THEN
        mask := 0;
        ph := 0.0;
        pm.Execute := TRUE;
        pm.N := 10;
        pm.CycleTime := 0.01;
        st := 1;
    END_IF;

    // drive DC samples: V=230, I=5 -> VRms~230, IRms~5, P~1150W, PF~1
    IF st = 1 THEN
        IF pm.Done THEN
            pm.Voltage := 230.0;
            pm.Current := 5.0;
            n := n + 1;
            IF n > 40 THEN
                IF pm.VRms > 140.0 THEN mask := mask + 1; END_IF;
                IF pm.IRms > 2.0 THEN mask := mask + 2; END_IF;
                IF pm.PReal > 200.0 THEN mask := mask + 4; END_IF;
                IF pm.PF > 0.8 THEN mask := mask + 8; END_IF;
                IF pm.Energy > 0.0 THEN mask := mask + 16; END_IF;
                st := 2;
            END_IF;
        END_IF;
    END_IF;

    pm();
END_PROGRAM

(* ---- tc2_qrc_case.st ---- *)
// tc2_qrc_case.st — QRC e2e: EAN-13 + UPC-A check-digit
// validation on known barcodes.
PROGRAM tc2_qrc_case
VAR
    q : FB_QrcValidate;
    st : INT;
    mask AT %QD0 : UDINT;
END_VAR
    IF st = 0 THEN
        mask := 0;
        q.Execute := TRUE;
        st := 1;
    ELSIF st = 1 THEN
        // EAN-13 5901234123457 — check digit 7
        q.D0 := 5; q.D1 := 9; q.D2 := 0; q.D3 := 1; q.D4 := 2;
        q.D5 := 3; q.D6 := 4; q.D7 := 1; q.D8 := 2; q.D9 := 3;
        q.D10 := 4; q.D11 := 5; q.D12 := 7;
        q.IsEan13 := TRUE;
        st := 2;
    ELSIF st = 2 THEN
        IF q.CodeOk THEN mask := mask + 1; END_IF;
        st := 3;
    ELSIF st = 3 THEN
        // EAN-13 wrong check — should be invalid
        q.D12 := 9;
        st := 4;
    ELSIF st = 4 THEN
        IF NOT q.CodeOk THEN mask := mask + 2; END_IF;
        st := 5;
    ELSIF st = 5 THEN
        // UPC-A 036000291452 — check digit 2
        q.D0 := 0; q.D1 := 3; q.D2 := 6; q.D3 := 0; q.D4 := 0;
        q.D5 := 0; q.D6 := 2; q.D7 := 9; q.D8 := 1; q.D9 := 4;
        q.D10 := 5; q.D11 := 2;
        q.IsEan13 := FALSE;
        st := 6;
    ELSIF st = 6 THEN
        IF q.CodeOk THEN mask := mask + 4; END_IF;
        st := 7;
    END_IF;

    q();
END_PROGRAM

(* ---- tc2_rfid_case.st ---- *)
// tc2_rfid_case.st — wired e2e for tc2_rfid (FB_RFIDReader).
PROGRAM tc2_rfid_case
VAR
    rd : FB_RFIDReader;
    st : INT;
    tries : INT;
    mask AT %QD0 : UDINT;
    diag AT %QD4 : UDINT;
END_VAR
    diag := st;
    IF st = 0 THEN
        mask := 0;
        rd.sDevice := '/tmp/rfid_pty';
        rd.nBaud := 9600; rd.nParity := 0;
        rd.nDataBits := 8; rd.nStopBits := 1;
        rd.sTxBuffer := 'READ';
        rd.nTxLen := 4;
        rd.tTimeout := T#500MS;
        rd.bExecute := TRUE;
        st := 1;
    ELSIF st = 1 THEN
        IF rd.bDone THEN mask := mask OR 1; END_IF;
        IF rd.hReader <> 0 THEN mask := mask OR 2; END_IF;
        IF rd.nRxLen > 0 THEN mask := mask OR 4; END_IF;
        IF FIND(rd.sRxBuffer, 'TAG:ABC12345') > 0 THEN
            mask := mask OR 8;
            rd.bExecute := FALSE;
            st := 2;
        ELSIF tries < 20 THEN
            // reader answers asynchronously: release, re-arm, retry
            tries := tries + 1;
            rd.bExecute := FALSE;
            st := 5;
        ELSE
            rd.bExecute := FALSE;
            st := 2;
        END_IF;
    ELSIF st = 5 THEN
        rd.bExecute := TRUE;                 // re-arm the cycle
        st := 6;
    ELSIF st = 6 THEN
        st := 1;
    ELSIF st = 2 THEN
        rd.bClose := TRUE;
        st := 3;
    ELSIF st = 3 THEN
        IF rd.hReader = 0 THEN mask := mask OR 16; END_IF;
        rd.bClose := FALSE;
        st := 4;
    END_IF;
    rd();
END_PROGRAM

(* ---- tc2_s5s7com_case.st ---- *)
PROGRAM Tc2S5S7ComCase
VAR
    mask      AT %QD0   : DINT;
    st        : INT;
    lnk       : FB_NLinkOpen;
    lnkBad    : FB_NLinkOpen;
    fch       : FB_NLinkFetch;
    fch2      : FB_NLinkFetch;
    fchBad    : FB_NLinkFetch;
    wr        : FB_NLinkWrite;
    wdata     : ARRAY[0..509] OF BYTE;
END_VAR

// autonomous S5 sequence against tests/compat/s5_test_peer.py
// (TCP 1103, RK512/3964). The peer serves DB1 (256B pattern
// (i*7+3)) and DB2 (256B pattern 0x40+(i&0x3F)). Each state's
// bExecute is high only while st equals its index, giving every
// FB one rising edge; bDone advances the machine.
wdata[0] := 16#DE; wdata[1] := 16#AD;
wdata[2] := 16#BE; wdata[3] := 16#EF;

lnk(sHost := '127.0.0.1', nPort := 1103, bExecute := st = 0,
    bClose := st = 9, tTimeout := T#3S);
lnkBad(sHost := '127.0.0.1', nPort := 19999, bExecute := st = 8,
       bClose := FALSE, tTimeout := T#3S);
fch(hLink := lnk.hLink, nArea := 1, nDB := 1, nOffset := 10,
    nLen := 16, bExecute := st = 1, tTimeout := T#2S);
wr(hLink := lnk.hLink, nArea := 1, nDB := 1, nOffset := 0,
   nLen := 4, pData := wdata, bExecute := st = 2,
   tTimeout := T#2S);
fch2(hLink := lnk.hLink, nArea := 1, nDB := 1, nOffset := 0,
     nLen := 4, bExecute := st = 3, tTimeout := T#2S);
fchBad(hLink := lnk.hLink, nArea := 1, nDB := 77, nOffset := 0,
       nLen := 4, bExecute := st = 4, tTimeout := T#2S);

IF st = 0 AND lnk.bDone THEN
    // connect -> READY, handle issued
    IF lnk.nStatus = 1 AND lnk.hLink <> 0 AND lnk.nErrID = 0 THEN
        mask := mask + 1;
    END_IF;
    st := 1;
ELSIF st = 1 AND fch.bDone THEN
    // DB1[10..25] = pattern (i*7+3): first byte 0x49, len 16
    IF fch.nStatus = 1 AND fch.cbRead = 16 AND fch.pBuffer[0] = 16#49
       AND fch.nErrID = 0 THEN
        mask := mask + 2;
    END_IF;
    st := 2;
ELSIF st = 2 AND wr.bDone THEN
    // SEND accepted
    IF wr.nStatus = 1 AND wr.cbWrite = 4 AND wr.nErrID = 0 THEN
        mask := mask + 4;
    END_IF;
    st := 3;
ELSIF st = 3 AND fch2.bDone THEN
    // read-back of the written bytes: wdata[0..3] = DE AD BE EF
    IF fch2.nStatus = 1 AND fch2.cbRead = 4
       AND fch2.pBuffer[0] = 16#DE AND fch2.pBuffer[1] = 16#AD
       AND fch2.pBuffer[2] = 16#BE AND fch2.pBuffer[3] = 16#EF
       AND fch2.nErrID = 0 THEN
        mask := mask + 8;
    END_IF;
    st := 4;
ELSIF st = 4 AND fchBad.bDone THEN
    // unknown DB -> RK512 status byte nonzero -> s5err
    IF fchBad.nStatus = 5 AND fchBad.nErrID <> 0 THEN
        mask := mask + 16;
    END_IF;
    st := 8;
ELSIF st = 8 AND lnkBad.bDone THEN
    // connect to a dead port -> conn error
    IF lnkBad.nStatus = 2 THEN
        mask := mask + 32;
    END_IF;
    st := 9;
ELSIF st = 9 AND lnk.bDone THEN
    st := 10;
END_IF;
END_PROGRAM

(* ---- tc2_serial_case.st ---- *)
PROGRAM Tc2SerialCase
VAR
    mask      AT %QD0   : DINT;
    st        : INT;
    scan_n    : UDINT;
    hPort     : UDINT;
    gotData   : STRING[256];
    gotLen    : UDINT;
    sentMsg   : STRING[256];
    open1     : FB_SerialOpen;
    openBad   : FB_SerialOpen;
    send1     : FB_SerialSend;
    recv1     : FB_SerialReceive;
    flush1    : FB_SerialFlush;
    rs485_1   : FB_SerialRs485;
    close1    : FB_SerialClose;
END_VAR

// autonomous pty loopback sequence: open -> send -> receive ->
// flush -> rs485 -> close, then a bad-path open for the error leg.
// sDevice is substituted by the test script with the pty slave path.
sentMsg := 'PING';

open1(bExecute := st = 0, tTimeout := T#5s,
      sDevice := '__PTY_SLAVE__', nBaud := 9600,
      nParity := 0, nDataBits := 8, nStopBits := 1, nFlags := 1);
openBad(bExecute := st = 5, tTimeout := T#5s,
        sDevice := '/nonexistent-tplc-serial', nBaud := 9600,
        nParity := 0, nDataBits := 8, nStopBits := 1, nFlags := 1);
send1(bExecute := st = 1, tTimeout := T#5s, hPort := hPort,
      pData := sentMsg, nLen := 4);
recv1(bExecute := st = 2, tTimeout := T#5s, hPort := hPort);
flush1(bExecute := st = 3, tTimeout := T#5s, hPort := hPort, nPurge := 3);
rs485_1(bExecute := st = 4, tTimeout := T#5s, hPort := hPort,
        bEnable := TRUE);
close1(bExecute := st = 5, tTimeout := T#5s, hPort := hPort);

IF st = 0 AND open1.bDone THEN
    IF open1.nErrId = 0 AND open1.hPort <> 0 THEN
        hPort := open1.hPort;
        mask := mask + 1;
    END_IF;
    st := 1;
ELSIF st = 1 AND send1.bDone THEN
    IF send1.nErrId = 0 AND send1.nSent = 4 THEN
        mask := mask + 2;
    END_IF;
    st := 2;
ELSIF st = 2 AND recv1.bDone THEN
    gotData := recv1.pData;
    gotLen := recv1.nRecBytes;
    IF recv1.nErrId = 0 AND recv1.nRecBytes = 4 THEN
        mask := mask + 4;
    END_IF;
    IF gotLen = 4 AND gotData = 'PING' THEN
        mask := mask + 8;
    END_IF;
    st := 3;
ELSIF st = 3 AND flush1.bDone THEN
    IF flush1.nErrId = 0 THEN
        mask := mask + 16;
    END_IF;
    st := 4;
ELSIF st = 4 AND rs485_1.bDone THEN
    IF rs485_1.nErrId = 0 THEN
        mask := mask + 32;
    END_IF;
    st := 5;
ELSIF st = 5 AND close1.bDone AND openBad.bDone THEN
    IF close1.nErrId = 0 AND openBad.nErrId = 3 THEN
        mask := mask + 64;
    END_IF;
    IF openBad.nErrId = 3 THEN
        mask := mask + 128;
    END_IF;
    st := 6;
END_IF;

scan_n := scan_n + 1;
END_PROGRAM

(* ---- tc2_sms_sms_case.st ---- *)
PROGRAM Tc2SmsSmtpCase
VAR
    mask      AT %QD0   : DINT;
    st        : INT;
    hPort     : UDINT;
    open1     : FB_SerialOpen;
    close1    : FB_SerialClose;
    sms1      : FB_SendSMS;
    smtp1     : FB_SmtpV3;
    smtp2     : FB_SmtpV3_Full;
    smtpBad   : FB_SmtpV3_Full;
    smtpDead  : FB_SmtpV3;
    attach1   : FB_SmtpAttach;
    ver1      : FB_GetTcPlcSMS_Version;
END_VAR

// autonomous sequence: open pty serial -> AT SMS -> SMTP plain
// -> SMTP auth -> SMTP reject -> attach-unsupported -> version
// -> refused connect -> close. sDevice is substituted by the
// test script with the pty slave path.

open1(bExecute := st = 0, tTimeout := T#5S,
      sDevice := '__PTY_SLAVE__', nBaud := 9600,
      nParity := 0, nDataBits := 8, nStopBits := 1, nFlags := 1);
close1(bExecute := st = 8, tTimeout := T#5S, hPort := hPort);

sms1(bExecute := st = 1, tTimeout := T#10S, hPort := hPort,
     sNumber := '+4915123456', sText := 'Hello TetherPLC');

smtp1(bExecute := st = 2, tTimeout := T#10S,
      sServer := '127.0.0.1', nPort := 2525,
      sFrom := 'plc@home.local', sTo := 'ops@example.com',
      sSubject := 'Plain Send',
      sBody := 'first line$N.second line dot-stuffed');

smtp2(bExecute := st = 3, tTimeout := T#10S,
      sServer := '127.0.0.1', nPort := 2525,
      sUser := 'alice', sPass := 's3cret',
      sFrom := 'plc@home.local', sTo := 'auth@example.com',
      sSubject := 'Auth Send', sBody := 'authenticated body');

smtpBad(bExecute := st = 4, tTimeout := T#10S,
        sServer := '127.0.0.1', nPort := 2525,
        sUser := 'alice', sPass := 's3cret',
        sFrom := 'plc@home.local', sTo := 'reject@example.com',
        sSubject := 'Reject', sBody := 'should fail');

attach1(bExecute := st = 5, tTimeout := T#10S,
        sServer := '127.0.0.1', nPort := 2525,
        sUser := '', sPass := '',
        sFrom := 'plc@home.local', sTo := 'ops@example.com',
        sSubject := 'Attach', sBody := 'x',
        sAttachPath := '/tmp/nope.bin');

ver1(bExecute := st = 6);

smtpDead(bExecute := st = 7, tTimeout := T#5S,
         sServer := '127.0.0.1', nPort := 2999,
         sFrom := 'plc@home.local', sTo := 'ops@example.com',
         sSubject := 'Dead', sBody := 'x');

IF st = 0 AND open1.bDone THEN
    IF open1.nErrId = 0 AND open1.hPort <> 0 THEN
        hPort := open1.hPort;
        mask := mask + 1;
    END_IF;
    st := 1;
ELSIF st = 1 AND sms1.bDone THEN
    IF sms1.nStatus = 0 AND sms1.bError = FALSE THEN
        mask := mask + 2;
    END_IF;
    st := 2;
ELSIF st = 2 AND smtp1.bDone THEN
    IF smtp1.nStatus = 1 AND smtp1.nRespCode = 250 THEN
        mask := mask + 4;
    END_IF;
    st := 3;
ELSIF st = 3 AND smtp2.bDone THEN
    IF smtp2.nStatus = 1 AND smtp2.nRespCode = 250 THEN
        mask := mask + 8;
    END_IF;
    st := 4;
ELSIF st = 4 AND smtpBad.bDone THEN
    IF smtpBad.nStatus = 2 AND smtpBad.nRespCode = 550 THEN
        mask := mask + 16;
    END_IF;
    st := 5;
ELSIF st = 5 AND attach1.bDone THEN
    IF attach1.nErrId = 90 AND attach1.bError THEN
        mask := mask + 32;
    END_IF;
    st := 6;
ELSIF st = 6 AND ver1.bDone THEN
    IF ver1.sVersion = 'TetherPLC-TcSMS 1.0' THEN
        mask := mask + 64;
    END_IF;
    st := 7;
ELSIF st = 7 AND smtpDead.bDone THEN
    IF smtpDead.nStatus >= 3 THEN
        mask := mask + 128;
    END_IF;
    st := 8;
ELSIF st = 8 AND close1.bDone THEN
    IF close1.nErrId = 0 THEN
        mask := mask + 256;
    END_IF;
    st := 9;
END_IF;

END_PROGRAM

(* ---- tc2_spa_case.st ---- *)
// tc2_spa_case.st — SPA e2e: peak detect, envelope, dft-bin,
// cross-correlation — pure-ST signal analysis.
PROGRAM tc2_spa_case
VAR
    pk : FB_PeakDetect;
    env : FB_Envelope;
    dft : FB_DftBin;
    xc : FB_XCorrQuality;
    st : INT;
    n : INT;
    mask AT %QD0 : UDINT;
    sig : LREAL;
END_VAR
    IF st = 0 THEN
        mask := 0;
        pk.Execute := TRUE;
        env.Execute := TRUE;
        dft.Execute := TRUE;
        xc.Execute := TRUE;
        pk.N := 8;
        env.AttackTn := 0.05; env.ReleaseTn := 0.5; env.CycleTime := 0.1;
        dft.N := 8; dft.Bin := 1; dft.CycleTime := 0.1;
        xc.N := 8;
        sig := 0.0;
        st := 1;
    END_IF;

    // drive a stepped signal
    IF st = 1 THEN
        n := n + 1;
        IF n < 4 THEN
            sig := 1.0;
        ELSIF n < 8 THEN
            sig := 4.0;   // peak
        ELSE
            sig := 2.0;
        END_IF;
        pk.Input := sig;
        env.Input := sig;
        dft.Input := sig;
        xc.Input := sig;
        xc.Reference := 2.0;
        IF n > 12 THEN
            IF pk.Peak >= 4.0 THEN mask := mask + 1; END_IF;   // saw peak
            IF pk.Valley <= 2.0 THEN mask := mask + 2; END_IF; // saw valley
            IF env.Output > 0.5 THEN mask := mask + 4; END_IF;  // envelope
            IF dft.Magnitude > 0.5 THEN mask := mask + 8; END_IF;
            st := 2;
        END_IF;
    END_IF;
    // cross-correlation of identical signals ~ +1
    IF st = 2 THEN
        n := n + 1;
        xc.Input := 2.0;
        xc.Reference := 2.0;
        IF n > 20 THEN
            IF xc.Quality > 0.9 THEN mask := mask + 16; END_IF; // ~+1
            st := 3;
        END_IF;
    END_IF;

    pk(); env(); dft(); xc();
END_PROGRAM

(* ---- tc2_system_ads_case.st ---- *)
PROGRAM Tc2SystemAdsCase
VAR
    mask      AT %QD0   : DINT;
    st        : INT;
    scan_n    : UDINT;
    hConn     : UDINT;
    gotData   : STRING[256];
    gotLen    : UDINT;
    wrData    : STRING[256];
    adsState  : DINT;
    devState  : DINT;
    conn1     : FB_AdsConnect;
    connBad   : FB_AdsConnect;
    read1     : FB_AdsRead;
    write1    : FB_AdsWrite;
    rstate1   : FB_AdsReadState;
    wctrl1    : FB_AdsWriteControl;
    bread1    : FB_AdsRead;
    close1    : FB_AdsClose;
END_VAR

// autonomous ADS exchange against the python test server:
// connect -> read -> write -> read-state -> write-control ->
// close, then a refused-port connect+read for the error leg.
wrData := 'WXYZ1234';

conn1(bExecute := st = 0, tTimeout := T#5s,
      sHost := '127.0.0.1', nPort := 18765);
connBad(bExecute := st = 5, tTimeout := T#5s,
        sHost := '127.0.0.1', nPort := 1);
read1(bExecute := st = 1, tTimeout := T#5s, hConn := hConn,
      nIdxGrp := 16#4020, nIdxOff := 0, nLen := 8);
write1(bExecute := st = 2, tTimeout := T#5s, hConn := hConn,
       nIdxGrp := 16#4020, nIdxOff := 8, pData := wrData, nLen := 8);
rstate1(bExecute := st = 3, tTimeout := T#5s, hConn := hConn);
wctrl1(bExecute := st = 4, tTimeout := T#5s, hConn := hConn,
       nAdsState := 5, nDevState := 0);
bread1(bExecute := st = 5 AND connBad.bDone, tTimeout := T#5s,
       hConn := connBad.hConn, nIdxGrp := 16#4020, nIdxOff := 0, nLen := 4);
close1(bExecute := st = 5, tTimeout := T#5s, hConn := hConn);

IF st = 0 AND conn1.bDone THEN
    IF conn1.nErrId = 0 AND conn1.hConn <> 0 THEN
        hConn := conn1.hConn;
        mask := mask + 1;
    END_IF;
    st := 1;
ELSIF st = 1 AND read1.bDone THEN
    gotData := read1.pData;
    gotLen := read1.nBytes;
    IF read1.nErrId = 0 AND read1.nAdsError = 0 AND
       read1.nBytes = 8 THEN
        mask := mask + 2;
    END_IF;
    IF gotLen = 8 AND gotData = 'ABCDEFGH' THEN
        mask := mask + 4;
    END_IF;
    st := 2;
ELSIF st = 2 AND write1.bDone THEN
    IF write1.nErrId = 0 AND write1.nAdsError = 0 THEN
        mask := mask + 8;
    END_IF;
    st := 3;
ELSIF st = 3 AND rstate1.bDone THEN
    adsState := rstate1.nAdsState;
    devState := rstate1.nDevState;
    IF rstate1.nErrId = 0 AND rstate1.nAdsError = 0 AND
       rstate1.nAdsState = 5 AND rstate1.nDevState = 0 THEN
        mask := mask + 16;
    END_IF;
    st := 4;
ELSIF st = 4 AND wctrl1.bDone THEN
    IF wctrl1.nErrId = 0 AND wctrl1.nAdsError = 0 THEN
        mask := mask + 32;
    END_IF;
    st := 5;
ELSIF st = 5 AND connBad.bDone AND bread1.bDone AND close1.bDone THEN
    IF close1.nErrId = 0 THEN
        mask := mask + 64;
    END_IF;
    IF bread1.nErrId = 3 THEN
        mask := mask + 128;
    END_IF;
    st := 6;
END_IF;

scan_n := scan_n + 1;
END_PROGRAM

(* ---- tc2_tc_case.st ---- *)
// tc2_tc_case.st — TempController e2e: a simulated thermal plant
// (heater -> PT1 lag -> sensor) driven by the PID+PWM controller.
PROGRAM tc2_tc_case
VAR
    ctl : FB_TempController;
    plant : LREAL;   // simulated thermal mass
    st : INT;
    n : INT;
    mask AT %QD0 : UDINT;
END_VAR
    IF st = 0 THEN
        mask := 0;
        plant := 20.0;                    // ambient
        ctl.Execute := TRUE;
        ctl.Setpoint := 100.0;
        ctl.Kp := 5.0; ctl.Tn := 1.0; ctl.Tv := 0.0;
        ctl.FilterTn := 0.5;
        ctl.PwmPeriod := 1.0;
        ctl.CycleTime := 0.1;
        st := 1;
    END_IF;

    // thermal plant: duty heats the mass, ambient cools it
    IF st = 1 THEN
        IF ctl.Done THEN
            n := n + 1;
            plant := plant +
                     (ctl.Duty * 0.02) - (plant - 20.0) * 0.001;
            ctl.Actual := plant;
            IF n > 50 THEN
                IF ctl.Duty > 10.0 THEN mask := mask + 1; END_IF;  // heating
                IF plant > 25.0 THEN mask := mask + 2; END_IF;     // rising
                IF ctl.Filtered > 20.0 THEN mask := mask + 4; END_IF;
                st := 2;
            END_IF;
        END_IF;
    END_IF;
    // keep driving — the plant settles toward SP
    IF st = 2 THEN
        IF ctl.Done THEN
            n := n + 1;
            plant := plant +
                     (ctl.Duty * 0.02) - (plant - 20.0) * 0.001;
            ctl.Actual := plant;
            IF n > 100 THEN
                IF plant > 30.0 THEN mask := mask + 8; END_IF;     // hot
                IF ctl.E < 90.0 THEN mask := mask + 16; END_IF;    // converging
                st := 3;
            END_IF;
        END_IF;
    END_IF;

    ctl();
END_PROGRAM

(* ---- tc2_tcpip_case.st ---- *)
PROGRAM Tc2TcpIpCase
VAR
    mask      AT %QD0   : DINT;
    st        : INT;
    scan_n    : UDINT;
    hListener : UDINT;
    hCli      : UDINT;
    hSrv      : UDINT;
    gotData   : STRING[256];
    gotLen    : UDINT;
    sentMsg   : STRING[256];
    listen1   : FB_SocketListen;
    conn1     : FB_SocketConnect;
    acc1      : FB_SocketAccept;
    send1     : FB_SocketSend;
    recv1     : FB_SocketReceive;
    closeCli  : FB_SocketClose;
    closeSrv  : FB_SocketClose;
    closeLst  : FB_SocketClose;
END_VAR

// autonomous loopback sequence: listen -> connect -> accept ->
// send -> receive -> close. Each state's bExecute is high only
// while st equals its index, giving every FB one rising edge.
sentMsg := 'PING';

listen1(bExecute := st = 0, tTimeout := T#5s,
        sHost := '', nPort := 17531);
conn1(bExecute := st = 1, tTimeout := T#5s,
      sHost := '127.0.0.1', nPort := 17531);
acc1(bExecute := st = 2, tTimeout := T#5s, hListener := hListener);
send1(bExecute := st = 3, tTimeout := T#5s, hSocket := hCli,
      pData := sentMsg, nLen := 4);
recv1(bExecute := st = 4, tTimeout := T#5s, hSocket := hSrv);
closeCli(bExecute := st = 5, tTimeout := T#5s, hSocket := hCli);
closeSrv(bExecute := st = 5, tTimeout := T#5s, hSocket := hSrv);
closeLst(bExecute := st = 5, tTimeout := T#5s, hSocket := hListener);

IF st = 0 AND listen1.bDone THEN
    IF listen1.nErrId = 0 AND listen1.hListener <> 0 THEN
        hListener := listen1.hListener;
        mask := mask + 1;
    END_IF;
    st := 1;
ELSIF st = 1 AND conn1.bDone THEN
    IF conn1.nErrId = 0 AND conn1.hSocket <> 0 THEN
        hCli := conn1.hSocket;
        mask := mask + 2;
    END_IF;
    st := 2;
ELSIF st = 2 AND acc1.bDone THEN
    IF acc1.bAccepted AND acc1.nErrId = 0 AND acc1.hSocket <> 0 THEN
        hSrv := acc1.hSocket;
        mask := mask + 4;
    END_IF;
    st := 3;
ELSIF st = 3 AND send1.bDone THEN
    IF send1.nErrId = 0 AND send1.nSent = 4 THEN
        mask := mask + 8;
    END_IF;
    st := 4;
ELSIF st = 4 AND recv1.bDone THEN
    gotData := recv1.pData;
    gotLen := recv1.nRecBytes;
    IF recv1.nErrId = 0 AND recv1.nRecBytes = 4 THEN
        mask := mask + 16;
    END_IF;
    IF gotLen = 4 AND gotData = 'PING' THEN
        mask := mask + 32;
    END_IF;
    st := 5;
ELSIF st = 5 AND closeCli.bDone AND closeSrv.bDone AND closeLst.bDone THEN
    IF closeCli.nErrId = 0 AND closeSrv.nErrId = 0 AND
       closeLst.nErrId = 0 THEN
        mask := mask + 64;
    END_IF;
    st := 6;
END_IF;

scan_n := scan_n + 1;
END_PROGRAM

(* ---- tc2_weighing_case.st ---- *)
// tc2_weighing_case.st — Weighing e2e: simulated load-cell signal,
// tare, net, stability, dosing coarse->fine->done.
PROGRAM tc2_weighing_case
VAR
    wgh : FB_Weigh;
    cell : LREAL;   // simulated load-cell signal
    st : INT;
    n : INT;
    mask AT %QD0 : UDINT;
END_VAR
    IF st = 0 THEN
        mask := 0;
        cell := 5.0;                      // empty cell = tare
        wgh.Execute := TRUE;
        wgh.FilterTn := 0.2;
        wgh.CycleTime := 0.1;
        wgh.DoTare := FALSE;              // tare captured in st=1
        wgh.StableBand := 0.05;
        wgh.StableCycles := 5;
        wgh.DoseSetpoint := 10.0;
        wgh.CoarseLimit := 0.8;
        st := 1;
    END_IF;

    // tare captured -> Net ~0
    IF st = 1 THEN
        IF wgh.Done THEN
            n := n + 1;
            cell := 5.0;                  // still empty
            wgh.Raw := cell;
            wgh.DoTare := TRUE;           // keep capturing tare
            IF n > 5 THEN
                IF wgh.TareWeight > 4.0 THEN mask := mask + 1; END_IF;
                IF wgh.Net < 1.0 THEN mask := mask + 2; END_IF;
                n := 0;
                wgh.DoTare := FALSE;
                st := 2;
            END_IF;
        END_IF;
    END_IF;
    // fill: cell signal ramps up
    IF st = 2 THEN
        IF wgh.Done THEN
            n := n + 1;
            cell := cell + 0.3;           // product filling
            wgh.Raw := cell;
            IF n > 30 THEN
                IF wgh.Net > 3.0 THEN mask := mask + 4; END_IF;
                n := 0;
                st := 3;
            END_IF;
        END_IF;
    END_IF;
    // dosing coarse->fine->done as Net approaches Setpoint
    IF st = 3 THEN
        IF wgh.Done THEN
            n := n + 1;
            cell := cell + 0.3;
            wgh.Raw := cell;
            IF wgh.DoseDone THEN
                mask := mask + 8;
                n := 0;
                st := 4;
            END_IF;
            IF n > 80 THEN st := 4; END_IF;
        END_IF;
    END_IF;
    // hold — verify stable flag settles
    IF st = 4 THEN
        IF wgh.Done THEN
            n := n + 1;
            IF n > 20 THEN
                IF wgh.Stable THEN mask := mask + 16; END_IF;
                st := 5;
            END_IF;
        END_IF;
    END_IF;

    wgh();
END_PROGRAM

(* ---- tc3_analytics_case.st ---- *)
// tc3_analytics_case.st — Tc3_Analytics e2e: counter+rate,
// windowed stats, ring logger, and honest engine-absent store.
PROGRAM tc3_analytics_case
VAR
    mask AT %QD0 : UDINT;
    cnt_ : FB_AnalyticsCounter;
    sts_ : FB_AnalyticsStats;
    lg_ : FB_AnalyticsLogger;
    sto_ : FB_AnalyticsStore;
    st : INT;
END_VAR
    // counter: 4 event edges in the first window, then rate>0
    IF st = 0 THEN
        mask := 0;
        cnt_.Enable := TRUE;
        cnt_.WindowTime := 0.05;
        cnt_.CycleTime := 0.01;
        cnt_.Event := FALSE;
        st := 1;
    ELSIF st = 1 THEN cnt_.Event := TRUE;  st := 2;
    ELSIF st = 2 THEN cnt_.Event := FALSE; st := 3;
    ELSIF st = 3 THEN cnt_.Event := TRUE;  st := 4;
    ELSIF st = 4 THEN cnt_.Event := FALSE; st := 5;
    ELSIF st = 5 THEN cnt_.Event := TRUE;  st := 6;
    ELSIF st = 6 THEN cnt_.Event := FALSE; st := 7;
    ELSIF st = 7 THEN cnt_.Event := TRUE;  st := 8;
    ELSIF st = 8 THEN
        cnt_.Event := FALSE;
        IF cnt_.Total = 4 THEN
            mask := mask OR 1;
            st := 9;
        END_IF;
    ELSIF st = 9 THEN
        IF cnt_.Rate > 0.0 THEN
            mask := mask OR 2;      // a window closed with events
            cnt_.Enable := FALSE;
            st := 10;
        END_IF;
    // stats: samples 2, 4, 9 -> count 3, min 2, max 9, mean 5
    ELSIF st = 10 THEN sts_.Execute := TRUE; sts_.Sample := 2.0; st := 11;
    ELSIF st = 11 THEN sts_.Sample := 4.0; st := 12;
    ELSIF st = 12 THEN sts_.Sample := 9.0; st := 13;
    ELSIF st = 13 THEN
        sts_.Execute := FALSE;
        IF sts_.Count = 3 AND sts_.Min = 2.0 AND sts_.Max = 9.0
           AND sts_.Mean > 4.9 AND sts_.Mean < 5.1 THEN
            mask := mask OR 4;
            st := 14;
        END_IF;
    // logger: 9 records -> wrap once, slot0 holds record 9
    ELSIF st = 14 THEN lg_.Record := TRUE;  lg_.Value := 10.0; lg_.Timestamp := 1.0; st := 15;
    ELSIF st = 15 THEN lg_.Record := FALSE; st := 16;
    ELSIF st = 16 THEN lg_.Record := TRUE;  lg_.Value := 20.0; lg_.Timestamp := 2.0; st := 17;
    ELSIF st = 17 THEN lg_.Record := FALSE; st := 18;
    ELSIF st = 18 THEN lg_.Record := TRUE;  lg_.Value := 30.0; lg_.Timestamp := 3.0; st := 19;
    ELSIF st = 19 THEN lg_.Record := FALSE; st := 20;
    ELSIF st = 20 THEN lg_.Record := TRUE;  lg_.Value := 40.0; lg_.Timestamp := 4.0; st := 21;
    ELSIF st = 21 THEN lg_.Record := FALSE; st := 22;
    ELSIF st = 22 THEN lg_.Record := TRUE;  lg_.Value := 50.0; lg_.Timestamp := 5.0; st := 23;
    ELSIF st = 23 THEN lg_.Record := FALSE; st := 24;
    ELSIF st = 24 THEN lg_.Record := TRUE;  lg_.Value := 60.0; lg_.Timestamp := 6.0; st := 25;
    ELSIF st = 25 THEN lg_.Record := FALSE; st := 26;
    ELSIF st = 26 THEN lg_.Record := TRUE;  lg_.Value := 70.0; lg_.Timestamp := 7.0; st := 27;
    ELSIF st = 27 THEN lg_.Record := FALSE; st := 28;
    ELSIF st = 28 THEN lg_.Record := TRUE;  lg_.Value := 80.0; lg_.Timestamp := 8.0; st := 29;
    ELSIF st = 29 THEN lg_.Record := FALSE; st := 30;
    ELSIF st = 30 THEN lg_.Record := TRUE;  lg_.Value := 90.0; lg_.Timestamp := 9.0; st := 31;
    ELSIF st = 31 THEN
        lg_.Record := FALSE;
        IF lg_.Count = 9 AND lg_.Overflow AND lg_.Slot0 = 90.0 AND lg_.LastTs = 9.0 THEN
            mask := mask OR 8;
            st := 32;
        END_IF;
    // store: provider configured -> honest engine-absent
    ELSIF st = 32 THEN
        sto_.ProviderPath := 'influx://db';
        sto_.RecordCount := 9;
        sto_.Execute := TRUE;
        st := 33;
    ELSIF st = 33 THEN
        IF sto_.Error AND sto_.ErrorId = 1 THEN
            mask := mask OR 16;
            st := 34;
        END_IF;
    ELSIF st = 34 THEN
        sto_.Execute := FALSE;
        st := 35;
    ELSIF st = 35 THEN
        sto_.ProviderPath := '';    // bad provider -> param error
        sto_.Execute := TRUE;
        st := 36;
    ELSIF st = 36 THEN
        IF sto_.Error AND sto_.ErrorId = 2 THEN
            mask := mask OR 32;
            st := 37;
        END_IF;
    END_IF;

    cnt_();
    sts_();
    lg_();
    sto_();
END_PROGRAM

(* ---- tc3_ba_common_case.st ---- *)
// tc3_ba_common_case.st — pure-ST e2e for tc3_ba_common.
PROGRAM tc3_ba_common_case
VAR
    rft : FB_BA_RFTrig;
    cov : FB_BA_ATrigCOV;
    rlm : FB_BA_RampLmt;
    sw2 : FB_BA_Swi2P;
    swh : FB_BA_SwiHys2P;
    pid : FB_BA_PIDCtrl;
    seq : FB_BA_SeqCtrl;
    arr : FB_BA_DynamicArray;
    rem : UDINT;
    okw : BOOL;
    st : INT;
    mask AT %QD0 : UDINT;
    zz : UDINT;
    diag AT %QD4 : UDINT;
END_VAR
    diag := st;
    mask := zz;
    IF st = 0 THEN
        zz := 0;
        pid.bEnable := TRUE;
        pid.fActual := 18.0; pid.fSetpoint := 22.0;
        pid.fKp := 2.0; pid.fTi := 0.0;
        pid.fOutMin := 0.0; pid.fOutMax := 100.0;
        pid.CycleTime := 0.1;
        rem := F_BA_RemSecsTp(10, 40);
        okw := F_BA_IsWeekdayValid(5);
        IF rem = 30 AND okw THEN zz := zz OR 1; END_IF;
        // COV trigger: first call reports
        cov.bEnable := TRUE;
        cov.fIn := 10.0;
        cov.fDelta := 1.0;
        st := 1;
    ELSIF st = 1 THEN
        IF pid.fOut > 5.0 THEN zz := zz OR 128; END_IF;
        IF cov.bTrig THEN zz := zz OR 2; END_IF;
        cov.fIn := 10.5;           // within delta: no trig
        st := 2;
    ELSIF st = 2 THEN
        IF NOT cov.bTrig THEN zz := zz OR 4; END_IF;
        cov.fIn := 12.5;           // delta 2.5: trig
        st := 3;
    ELSIF st = 3 THEN
        IF cov.bTrig THEN zz := zz OR 8; END_IF;
        // ramp limiter
        rlm.bEnable := TRUE;
        rlm.fIn := 50.0; rlm.fSlewUp := 10.0; rlm.fSlewDown := 10.0;
        rlm.fMin := 0.0; rlm.fMax := 40.0;
        rlm.CycleTime := 0.1;
        st := 4;
    ELSIF st = 4 THEN
        IF rlm.fOut = 40.0 THEN zz := zz OR 16; st := 5; END_IF;
        IF rlm.fOut > 40.0 THEN diag := 16#E4; st := 99; END_IF;
    ELSIF st = 5 THEN
        // switches
        sw2.bEnable := TRUE;
        sw2.fIn := 6.0; sw2.fOn := 5.0; sw2.fOff := 1.0;
        swh.bEnable := TRUE;
        swh.fIn := 18.0; swh.fSp := 21.0; swh.fHys := 2.0;
        swh.bInvert := FALSE;      // heating: on below SP-hys
        st := 6;
    ELSIF st = 6 THEN
        IF sw2.bOut THEN zz := zz OR 32; END_IF;
        IF swh.bOut THEN zz := zz OR 64; END_IF;
        // PID
        // seq: demand 60 across 3 stages -> s1 100, s2 80, s3 0
        seq.bEnable := TRUE;
        seq.fDemand := 60.0; seq.nStages := 3;
        st := 7;
    ELSIF st = 7 THEN
        st := 20;
    ELSIF st = 20 THEN
        IF seq.fStage1 > 99.0 AND seq.fStage2 > 75.0 AND
           seq.fStage2 < 85.0 AND seq.fStage3 < 1.0 THEN
            zz := zz OR 256;
        END_IF;
        // dynamic array: set/get/remove
        arr.bEnable := TRUE;
        arr.Op := 1;               // set
        arr.Key := 7;
        arr.Value := 42.0;
        st := 8;
    ELSIF st = 8 THEN
        IF arr.Done THEN zz := zz OR 512; END_IF;
        arr.Op := 2;               // get
        arr.Key := 7;
        st := 9;
    ELSIF st = 9 THEN
        IF arr.Found AND arr.OutValue = 42.0 THEN zz := zz OR 1024; END_IF;
        arr.Op := 3;               // remove
        arr.Key := 7;
        st := 10;
    ELSIF st = 10 THEN
        IF arr.Done THEN zz := zz OR 2048; END_IF;
        arr.Op := 4;               // find (should miss)
        arr.Key := 7;
        st := 11;
    ELSIF st = 11 THEN
        IF NOT arr.Found THEN zz := zz OR 4096; END_IF;
        arr.Op := 0;
        // edge trigger
        rft.bIn := TRUE;
        st := 12;
    ELSIF st = 12 THEN
        IF rft.bRise THEN zz := zz OR 8192; END_IF;
        rft.bIn := FALSE;
        st := 13;
    ELSIF st = 13 THEN
        IF rft.bFall THEN zz := zz OR 16384; END_IF;
        st := 14;
    END_IF;

    rft(); cov(); rlm(); sw2(); swh(); pid(); seq(); arr();
END_PROGRAM

(* ---- tc3_bacnet_case.st ---- *)
PROGRAM Tc3BacnetCase
VAR
    mask      AT %QD0   : DINT;
    st        : INT;
    w         : FB_BACnet_WhoIs;
    w2        : FB_BACnet_WhoIs;
    r         : FB_BACnet_ReadProperty;
    wr        : FB_BACnet_WriteProperty;
    rn        : FB_BACnet_ReadProperty;
    re        : FB_BACnet_ReadProperty;
    wval      : ARRAY[0..255] OF BYTE;
END_VAR

// autonomous BACnet/IP sequence against tests/compat/
// bacnet_test_peer.py (UDP 47808): broadcast Who-Is with a
// 1000..2000 instance range -> I-Am; ReadProperty real /
// unsigned / object-name; WriteProperty Simple-ACK; Error for
// the unknown object. Each state's bExecute is high only while
// st equals its index, giving every FB one rising edge.
wval[0] := 16#41;
wval[1] := 16#64;
wval[2] := 16#00;
wval[3] := 16#00;   // REAL 22.5 big-endian payload

w(bExecute := st = 0, sHost := '255.255.255.255', nPort := 47808,
  bHasRange := TRUE, nRangeLo := 1000, nRangeHi := 2000,
  tTimeout := T#1S);
r(bExecute := st = 1, sHost := '127.0.0.1', nPort := 47808,
  nObjType := 0, nObjInst := 1, nPropId := 85,
  bHasIdx := FALSE, nPropIdx := 0, tTimeout := T#1S);
wr(bExecute := st = 2, sHost := '127.0.0.1', nPort := 47808,
   nObjType := 1, nObjInst := 1, nPropId := 85,
   bHasIdx := FALSE, nPropIdx := 0,
   nValueType := 4, nValueLen := 4, pValue := wval,
   bHasPrio := TRUE, nPriority := 8, tTimeout := T#1S);
rn(bExecute := st = 3, sHost := '127.0.0.1', nPort := 47808,
   nObjType := 8, nObjInst := 1234, nPropId := 77,
   bHasIdx := FALSE, nPropIdx := 0, tTimeout := T#1S);
re(bExecute := st = 4, sHost := '127.0.0.1', nPort := 47808,
   nObjType := 0, nObjInst := 9999, nPropId := 85,
   bHasIdx := FALSE, nPropIdx := 0, tTimeout := T#1S);
w2(bExecute := st = 5, sHost := '127.0.0.1', nPort := 47808,
   bHasRange := FALSE, nRangeLo := 0, nRangeHi := 0,
   tTimeout := T#1S);

IF st = 0 AND w.bDone THEN
    // broadcast I-Am: device(8).1234, vendor 260, maxAPDU 1476,
    // segmentation 0; the reply source is the routed interface
    // address, so only check that dev_ip was populated
    IF w.nDevCount >= 1 AND w.nDevId[0] = 33555666 AND
       NOT (w.nDevIp[0] = 0 AND w.nDevIp[1] = 0 AND
            w.nDevIp[2] = 0 AND w.nDevIp[3] = 0) AND
       w.nDevVendor = 260 AND w.nDevMaxApdu = 1476 AND
       w.nDevSeg = 0 AND w.nErrId = 0 THEN
        mask := mask + 1;
    END_IF;
    st := 1;
ELSIF st = 1 AND r.bDone THEN
    // Complex-ACK echoes obj/prop; value = REAL 21.5 (41 AC 00 00)
    IF r.nStatus = 1 AND r.nService = 12 AND r.nValueType = 4 AND
       r.nValueLen = 4 AND r.pValue[0] = 16#41 AND
       r.pValue[1] = 16#AC AND r.pValue[2] = 16#00 AND
       r.pValue[3] = 16#00 AND r.nRObjType = 0 AND
       r.nRObjInst = 1 AND r.nRPropId = 85 AND r.nErrId = 0 THEN
        mask := mask + 2;
    END_IF;
    st := 2;
ELSIF st = 2 AND wr.bDone THEN
    IF wr.nStatus = 1 AND wr.nService = 15 AND wr.nErrId = 0 THEN
        mask := mask + 4;
    END_IF;
    st := 3;
ELSIF st = 3 AND rn.bDone THEN
    // object-name 'TETH-PLC' = 54 45 54 48 2D 50 4C 43
    IF rn.nStatus = 1 AND rn.nValueType = 7 AND rn.nValueLen = 8 AND
       rn.pValue[0] = 16#54 AND rn.pValue[1] = 16#45 AND
       rn.pValue[4] = 16#2D AND rn.pValue[7] = 16#43 AND
       rn.nRObjType = 8 AND rn.nRObjInst = 1234 AND
       rn.nRPropId = 77 AND rn.nErrId = 0 THEN
        mask := mask + 8;
    END_IF;
    st := 4;
ELSIF st = 4 AND re.bDone THEN
    // unknown object -> BACnet Error APDU -> STATUS 3
    IF re.nStatus = 3 AND re.nErrId = 0 THEN
        mask := mask + 16;
    END_IF;
    st := 5;
ELSIF st = 5 AND w2.bDone THEN
    // directed (BVLC unicast) Who-Is: reply source is 127.0.0.1
    IF w2.nDevCount >= 1 AND w2.nDevId[0] = 33555666 AND
       w2.nDevIp[0] = 127 AND w2.nDevIp[1] = 0 AND
       w2.nDevIp[2] = 0 AND w2.nDevIp[3] = 1 AND w2.nErrId = 0 THEN
        mask := mask + 32;
    END_IF;
    st := 6;
END_IF;

END_PROGRAM

(* ---- tc3_database_case.st ---- *)
// tc3_database_case.st — e2e for tc3_database (tplc-db/SQLite).
PROGRAM tc3_database_case
VAR
    opn : FB_PLCDBOpen;
    ddl : FB_PLCDBCreateEvt;
    wr1 : FB_PLCDBWriteEvt;
    wr2 : FB_PLCDBWriteEvt;
    rd : FB_PLCDBReadEvt;
    er : FB_PLCDBGetError;
    st : INT;
    mask AT %QD0 : UDINT;
    diag AT %QD4 : UDINT;
END_VAR
    diag := st;
    IF st = 0 THEN
        mask := 0;
        opn.sPath := '/tmp/tplc_db_e2e.sqlite';
        opn.nCmd := 1;
        st := 1;
    ELSIF st = 1 THEN
        IF opn.bDone AND opn.hDb <> 0 THEN mask := mask OR 1; END_IF;
        opn.nCmd := 0;
        ddl.hDb := opn.hDb;
        ddl.sSql := 'CREATE TABLE IF NOT EXISTS tags (id INTEGER, val INTEGER)';
        st := 2;
    ELSIF st = 2 THEN
        ddl.nCmd := 2;
        st := 3;
    ELSIF st = 3 THEN
        IF ddl.bDone THEN mask := mask OR 2; END_IF;
        ddl.nCmd := 0;
        wr1.hDb := opn.hDb;
        wr1.sSql := 'DELETE FROM tags';
        st := 4;
    ELSIF st = 4 THEN
        wr1.nCmd := 2;
        st := 5;
    ELSIF st = 5 THEN
        IF wr1.bDone THEN mask := mask OR 4; END_IF;
        wr1.nCmd := 0;
        wr2.hDb := opn.hDb;
        wr2.sSql := 'INSERT INTO tags VALUES (2, 21), (1, 7)';
        st := 6;
    ELSIF st = 6 THEN
        wr2.nCmd := 2;
        st := 7;
    ELSIF st = 7 THEN
        IF wr2.bDone AND wr2.nChanges = 2 THEN mask := mask OR 8; END_IF;
        wr2.nCmd := 0;
        rd.hDb := opn.hDb;
        rd.sSql := 'SELECT id, val FROM tags ORDER BY id';
        st := 8;
    ELSIF st = 8 THEN
        rd.nCmd := 3;
        st := 9;
    ELSIF st = 9 THEN
        IF rd.bDone AND rd.nRows = 2 AND rd.nCols = 2 THEN
            mask := mask OR 16;
        END_IF;
        // rows: "1\t7\n2\t21\n"
        IF FIND(rd.sResult, '1') = 1 THEN mask := mask OR 32; END_IF;
        IF FIND(rd.sResult, '21') > 0 THEN mask := mask OR 64; END_IF;
        IF FIND(rd.sResult, '21') > 0 THEN mask := mask OR 128; END_IF;
        rd.nCmd := 0;
        rd.sSql := 'SELECT nope FROM tags';
        st := 10;
    ELSIF st = 10 THEN
        rd.nCmd := 3;                        // bad SQL -> error
        st := 11;
    ELSIF st = 11 THEN
        IF rd.bError THEN mask := mask OR 256; END_IF;
        rd.nCmd := 0;
        er.hDb := opn.hDb;
        st := 12;
    ELSIF st = 12 THEN
        er.nCmd := 5;                        // engine error text
        st := 13;
    ELSIF st = 13 THEN
        IF er.bDone AND FIND(er.sError, 'nope') > 0 THEN
            mask := mask OR 512;
        END_IF;
        er.nCmd := 0;
        opn.nCmd := 4;                       // close
        st := 14;
    ELSIF st = 14 THEN
        IF opn.bDone AND opn.hDb = 0 THEN mask := mask OR 1024; END_IF;
        opn.nCmd := 0;
        st := 15;
    END_IF;
    opn(); ddl(); wr1(); wr2(); rd(); er();
END_PROGRAM

(* ---- tc3_dynmem_case.st ---- *)
// tc3_dynmem_case.st — e2e for tc3_dynmem (tplc-dynmem arena).
// Convention: a state that sets nCmd executes at that scan's
// FB call; the next state checks *Done and clears nCmd so the
// following command sees a fresh edge.
PROGRAM tc3_dynmem_case
VAR
    buf : FB_DynMem_Buffer;
    acc : FB_DynMem_Access;
    mgr : FB_DynMem_Manager;
    st : INT;
    mask AT %QD0 : UDINT;
    diag AT %QD4 : UDINT;
END_VAR
    diag := st;
    IF st = 0 THEN
        mask := 0;
        buf.bReset := TRUE;
        buf.nNewSize := 16; buf.nCmd := 1;   // alloc 16, zeroed
        st := 1;
    ELSIF st = 1 THEN
        IF buf.bDone AND buf.hBuffer <> 0 THEN mask := mask OR 1; END_IF;
        buf.nCmd := 0;
        acc.nHandle := buf.hBuffer; acc.nOffset := 3;
        acc.nByte := 16#A5;
        st := 2;
    ELSIF st = 2 THEN
        acc.nCmd := 5;                       // write 0xA5@3
        st := 3;
    ELSIF st = 3 THEN
        IF acc.bDone THEN mask := mask OR 2; END_IF;
        acc.nCmd := 0;
        st := 4;
    ELSIF st = 4 THEN
        acc.nCmd := 4;                       // read it back
        st := 5;
    ELSIF st = 5 THEN
        IF acc.bDone AND acc.nOut = 16#A5 THEN mask := mask OR 4; END_IF;
        acc.nCmd := 0;
        buf.bPreserve := TRUE; buf.bReset := FALSE;
        buf.nNewSize := 32;
        st := 6;
    ELSIF st = 6 THEN
        buf.nCmd := 2;                       // realloc grow, preserve
        st := 7;
    ELSIF st = 7 THEN
        IF buf.bDone AND buf.nSize = 32 THEN mask := mask OR 8; END_IF;
        buf.nCmd := 0;
        st := 8;
    ELSIF st = 8 THEN
        acc.nHandle := buf.hBuffer; acc.nOffset := 3;
        acc.nCmd := 4;                       // preserved byte?
        st := 9;
    ELSIF st = 9 THEN
        IF acc.bDone AND acc.nOut = 16#A5 THEN mask := mask OR 16; END_IF;
        acc.nCmd := 0;
        acc.nOffset := 64;
        st := 10;
    ELSIF st = 10 THEN
        acc.nCmd := 4;                       // out-of-range -> error
        st := 11;
    ELSIF st = 11 THEN
        IF acc.bError THEN mask := mask OR 32; END_IF;
        acc.nCmd := 0;
        st := 12;
    ELSIF st = 12 THEN
        buf.nCmd := 3;                       // deallocate
        st := 13;
    ELSIF st = 13 THEN
        IF buf.bDone AND buf.hBuffer = 0 THEN mask := mask OR 64; END_IF;
        buf.nCmd := 0;
        mgr.nReqSize := 8;
        st := 14;
    ELSIF st = 14 THEN
        mgr.nCmd := 1;                       // manager alloc
        st := 15;
    ELSIF st = 15 THEN
        IF mgr.bDone AND mgr.hNew <> 0
           AND mgr.nLiveBlocks = 1 AND mgr.nLiveBytes = 8 THEN
            mask := mask OR 128;
        END_IF;
        mgr.nCmd := 0;
        mgr.nId := mgr.hNew;
        st := 16;
    ELSIF st = 16 THEN
        mgr.nCmd := 3;                       // manager dealloc
        st := 17;
    ELSIF st = 17 THEN
        IF mgr.bDone AND mgr.nLiveBlocks = 0
           AND mgr.nTotalFrees = 2 THEN
            mask := mask OR 256;
        END_IF;
        mgr.nCmd := 0;
        st := 18;
    END_IF;
    buf(); acc(); mgr();
END_PROGRAM

(* ---- tc3_ecdiag_case.st ---- *)
// tc3_ecdiag_case.st — Tc3_EtherCATDiag e2e against
// tether_io_motion_server (TPLC_EC_IO): read the simulated CoE
// 0x10F3 diag history for slave 0 (3 entries: info/warning/error),
// verify decoded fields, acknowledge, re-read, then check slave 1
// (2 entries) and slave 5 (empty).  ELSIF chain prevents same-scan
// state cascade.
PROGRAM tc3_ecdiag_case
VAR
    rd : FB_CoE_DiagHistory_Read;
    st : INT;
    waitN : INT;
    mask AT %QD0 : UDINT;
    ok1 : BOOL;
    ok2 : BOOL;
    ok3 : BOOL;
    ok4 : BOOL;
    ok5 : BOOL;
    ok6 : BOOL;
    ok7 : BOOL;
    ok8 : BOOL;
    ok9 : BOOL;
END_VAR
    IF st = 0 THEN
        mask := 0;
        waitN := 0;
        rd.nSlaveAddr := 0;
        rd.bEnable := TRUE;
        rd.bAck := FALSE;
        rd.nReadIntervalScans := 100000;
        st := 1;
    ELSIF st = 1 THEN
        // first read complete when bValid or bError
        IF rd.bValid OR rd.bError THEN
            ok1 := rd.oCount = 3 AND rd.oNewest = 3 AND
                    rd.oAcked = 2 AND rd.oNewMsgs = 1 AND
                    NOT rd.bError;
            IF ok1 THEN mask := mask + 1; END_IF;
            ok2 := rd.aEMsgType[0] = 1 AND rd.aEMsgType[1] = 2 AND
                    rd.aEMsgType[2] = 3;
            IF ok2 THEN mask := mask + 2; END_IF;
            ok3 := rd.aEAckStatus[0] = 1 AND rd.aEAckStatus[1] = 1 AND
                    rd.aEAckStatus[2] = 0;
            IF ok3 THEN mask := mask + 4; END_IF;
            ok4 := rd.aEDiagCode[0] = 16#1000 AND
                    rd.aEDiagCode[1] = 16#1001 AND
                    rd.aEDiagCode[2] = 16#E0008105 AND
                    rd.aETextId[0] = 16#1100 AND
                    rd.aETextId[2] = 16#8105;
            IF ok4 THEN mask := mask + 8; END_IF;
            ok5 := rd.aEModuleNo[2] = 1 AND rd.aEChannelNo[2] = 2 AND
                    rd.aEDiagCodeType[2] = 3;
            IF ok5 THEN mask := mask + 16; END_IF;
            ok6 := rd.aETimestampMs[0] = 1000 AND
                    rd.aETimestampMs[1] = 2000 AND
                    rd.aETimestampMs[2] = 3000;
            IF ok6 THEN mask := mask + 32; END_IF;
            rd.bAck := TRUE;
            st := 2;
        ELSIF waitN > 60 THEN
            st := 90;
        ELSE
            waitN := waitN + 1;
        END_IF;
    ELSIF st = 2 THEN
        // ack edge consumed; wait for the post-ack read
        IF rd.bValid OR rd.bError THEN
            ok7 := rd.oAcked = 3 AND rd.oNewMsgs = 0 AND
                    rd.aEAckStatus[0] = 1 AND rd.aEAckStatus[1] = 1 AND
                    rd.aEAckStatus[2] = 1;
            IF ok7 THEN mask := mask + 64; END_IF;
            rd.bAck := FALSE;
            rd.bEnable := FALSE;
            rd.nSlaveAddr := 1;
            waitN := 0;
            st := 3;
        ELSIF waitN > 60 THEN
            st := 90;
        ELSE
            waitN := waitN + 1;
        END_IF;
    ELSIF st = 3 THEN
        rd.bEnable := TRUE;   // rising edge -> read slave 1
        st := 4;
    ELSIF st = 4 THEN
        IF rd.bValid OR rd.bError THEN
            ok8 := rd.oCount = 2 AND rd.oNewest = 2;
            IF ok8 THEN mask := mask + 128; END_IF;
            rd.bEnable := FALSE;
            rd.nSlaveAddr := 5;
            waitN := 0;
            st := 5;
        ELSIF waitN > 60 THEN
            st := 90;
        ELSE
            waitN := waitN + 1;
        END_IF;
    ELSIF st = 5 THEN
        rd.bEnable := TRUE;
        st := 6;
    ELSIF st = 6 THEN
        IF rd.bValid OR rd.bError THEN
            ok9 := rd.oCount = 0 AND rd.oNewest = 0 AND
                    NOT rd.bError;
            IF ok9 THEN mask := mask + 256; END_IF;
            rd.bEnable := FALSE;
            st := 90;
        ELSIF waitN > 60 THEN
            st := 90;
        ELSE
            waitN := waitN + 1;
        END_IF;
    ELSIF st = 90 THEN
        // done; mask holds results
    END_IF
    rd();
END_PROGRAM

(* ---- tc3_ecsync_case.st ---- *)
// tc3_ecsync_case.st — Tc3_EtherCATExtSync e2e against
// tether_io_motion_server (TPLC_EC_IO): enable sync -> TS1Done,
// windowed IsSynchronized checks, disable, re-enable.
// ELSIF chain prevents same-scan state cascade; each state does one
// thing per scan.
PROGRAM tc3_ecsync_case
VAR
    ext : FB_EcExtSyncExtTimes;
    iso : FB_EcExtSyncIsSynchronized;
    st : INT;
    waitN : INT;
    mask AT %QD0 : UDINT;
    netid : STRING[22];
    sBig : BOOL;
    ncBig : BOOL;
    sNarrow : BOOL;
    ncNarrow : BOOL;
    sOff : BOOL;
    ncOff : BOOL;
END_VAR
    IF st = 0 THEN
        mask := 0;
        netid := '';
        waitN := 0;
        st := 1;
    ELSIF st = 1 THEN
        netid := '1.2.3.4:5.6';
        st := 2;
    ELSIF st = 2 THEN
        IF ext.bTS1Done THEN
            IF NOT ext.bError THEN mask := mask + 1; END_IF;
            st := 3;
        ELSIF waitN > 60 THEN
            st := 90;   // timeout -> fail state
        ELSE
            waitN := waitN + 1;
        END_IF;
    ELSIF st = 3 THEN
        iso.nSyncWindow := 4000000000;
        iso();
        sBig := iso.bSynchronized;
        ncBig := iso.bNotConnected;
        iso.nSyncWindow := 500;
        iso();
        sNarrow := iso.bSynchronized;
        ncNarrow := iso.bNotConnected;
        IF sBig AND NOT ncBig AND NOT ncNarrow AND NOT sNarrow
           AND NOT iso.bError THEN
            mask := mask + 2;
        END_IF;
        netid := '';
        st := 4;
    ELSIF st = 4 THEN
        // sync disabled: neither synchronized nor not-connected
        iso.nSyncWindow := 4000000000;
        iso();
        sOff := iso.bSynchronized;
        ncOff := iso.bNotConnected;
        IF NOT sOff AND NOT ncOff AND NOT iso.bError THEN
            mask := mask + 4;
        END_IF;
        netid := '1.2.3.4:5.6';
        waitN := 0;
        st := 5;
    ELSIF st = 5 THEN
        IF ext.bTS1Done THEN
            iso.nSyncWindow := 4000000000;
            iso();
            IF iso.bSynchronized AND NOT iso.bNotConnected THEN
                mask := mask + 8;
            END_IF;
            st := 6;
        ELSIF waitN > 60 THEN
            st := 90;
        ELSE
            waitN := waitN + 1;
        END_IF;
    ELSIF st = 6 THEN
        st := 90;
    ELSIF st = 90 THEN
        // done; mask holds results
    END_IF
    ext.sNetId := netid;
    ext();
    iso();
END_PROGRAM

(* ---- tc3_ecsync_nosvc_case.st ---- *)
// tc3_ecsync_nosvc_case.st — negative e2e: no TPLC_EC_IO endpoint,
// so tplc-ecsync is inactive and both FBs must report the link as
// not connected with a service error.
PROGRAM tc3_ecsync_nosvc_case
VAR
    ext : FB_EcExtSyncExtTimes;
    iso : FB_EcExtSyncIsSynchronized;
    st : INT;
    mask AT %QD0 : UDINT;
    netid : STRING[22];
END_VAR
    IF st = 0 THEN
        mask := 0;
        netid := '';
        iso.nSyncWindow := 4000000000;
        st := 1;
    ELSIF st = 1 THEN
        iso();
        IF iso.bNotConnected AND iso.bError AND NOT iso.bSynchronized THEN
            mask := mask + 1;
        END_IF;
        netid := '1.2.3.4:5.6';
        st := 2;
    ELSIF st = 2 THEN
        IF ext.bError AND NOT ext.bTS1Done THEN
            mask := mask + 2;
        END_IF;
        st := 3;
    ELSIF st = 3 THEN
        // hold
    END_IF
    ext.sNetId := netid;
    ext();
    iso();
END_PROGRAM
